// get enumerations from XPU for visu:	
GVL_APPLICATION.VisuPoolData.eTransportState                       := f_GetState   (GVL_XTS.XtsTransportState.State);
GVL_APPLICATION.VisuPoolData.eTransportResult                      := f_GetProgress(GVL_XTS.XtsTransportState.State);
GVL_APPLICATION.VisuPoolData.eXpuState                             := f_GetState   (GVL_XTS.XtsTransportState.XpuState.State);
GVL_APPLICATION.VisuPoolData.eXpuResult                            := f_GetProgress(GVL_XTS.XtsTransportState.XpuState.State);
GVL_APPLICATION.VisuPoolData.eXpuCheck                             := GVL_XTS.XtsTransportState.XpuState.Check;

// display xpu state and result in visu
// get strings and info
GVL_APPLICATION.VisuPoolData.sCaGroupState                         := TO_STRING(GVL_XTS.XtsTransportState.GroupInfo.CaGroupState);

GVL_APPLICATION.VisuPoolData.sTransportState                       := TO_STRING(GVL_APPLICATION.VisuPoolData.eTransportState);
GVL_APPLICATION.VisuPoolData.sTransportCheck                       := TO_STRING(GVL_XTS.XtsTransportState.Check);
GVL_APPLICATION.VisuPoolData.sTransportResult                      := TO_STRING(GVL_APPLICATION.VisuPoolData.eTransportResult);

GVL_APPLICATION.VisuPoolData.stXpuStrings.sXpuState                := TO_STRING(GVL_APPLICATION.VisuPoolData.eXpuState);
GVL_APPLICATION.VisuPoolData.stXpuStrings.sXpuResult               := TO_STRING(GVL_APPLICATION.VisuPoolData.eXpuResult);
GVL_APPLICATION.VisuPoolData.stXpuStrings.sXpuCyclicCheck          := TO_STRING(GVL_APPLICATION.VisuPoolData.eXpuCheck);

GVL_APPLICATION.VisuPoolData.stXpuStrings.sXpuOpMode               := TO_STRING(GVL_XTS.XtsTransportState.XpuInfo.OperationMode);
GVL_APPLICATION.VisuPoolData.stXpuStrings.sXpuMoverId_DetectionMode:= TO_STRING(GVL_XTS.XtsTransportState.XpuInfo.IdDetectionMode);
GVL_APPLICATION.VisuPoolData.stXpuStrings.sXpuMoverPosAssignement  := TO_STRING(GVL_XTS.XtsTransportState.XpuInfo.MoverPositionAssignement);
//---------------------------------------------------------------------------------------------------------------
// check the indices before access
//---------------------------------------------------------------------------------------------------------------
nMoverSelected       := SEL((nMoverSelected<1),                               nMoverSelected, 1);
nMoverSelected       := SEL((nMoverSelected>GVL_XTS_CONSTANTS.MAX_MOVER),     nMoverSelected, GVL_XTS_CONSTANTS.MAX_MOVER);

nStationSelected     := SEL((nStationSelected<1),                             nStationSelected, 1);
nStationSelected     := SEL((nStationSelected>GVL_XTS_CONSTANTS.MAX_STATION), nStationSelected, GVL_XTS_CONSTANTS.MAX_STATION);

nCollectorSelected   := SEL((nCollectorSelected<1),                           nCollectorSelected, 1);
nCollectorSelected   := SEL((nCollectorSelected>GVL_APPLICATION.MAX_PROCESS), nCollectorSelected, GVL_APPLICATION.MAX_PROCESS);

nInstanceSelected    := SEL((nInstanceSelected<1),                            nInstanceSelected, 1);
nInstanceSelected    := SEL((nInstanceSelected>GVL_APPLICATION.MAX_PROCESS),  nInstanceSelected, GVL_APPLICATION.MAX_PROCESS);
//---------------------------------------------------------------------------------------------------------------
// get indexed data
//---------------------------------------------------------------------------------------------------------------
GVL_APPLICATION.VisuPoolData.eMoverState        := f_GetState   (GVL_XTS.MoverState[nMoverSelected].State);
GVL_APPLICATION.VisuPoolData.eMoverResult       := f_GetProgress(GVL_XTS.MoverState[nMoverSelected].State);
GVL_APPLICATION.VisuPoolData.sMoverState        := TO_STRING(GVL_APPLICATION.VisuPoolData.eMoverState);
GVL_APPLICATION.VisuPoolData.sMoverResult       := TO_STRING(GVL_APPLICATION.VisuPoolData.eMoverResult);

GVL_APPLICATION.VisuPoolData.bStationEnable     := SEL((GVL_XTS.StationCtrl[nStationSelected].Cmd = E_STATION_CTRL.STATION_ENABLE),        FALSE, TRUE);
GVL_APPLICATION.VisuPoolData.bStationEnter      := SEL((GVL_XTS.StationCtrl[nStationSelected].Cmd = E_STATION_CTRL.STATION_MOVER_ENTER),   FALSE, TRUE);
GVL_APPLICATION.VisuPoolData.bStationStart      := SEL((GVL_XTS.StationCtrl[nStationSelected].Cmd = E_STATION_CTRL.STATION_PROCESS_START), FALSE, TRUE);
GVL_APPLICATION.VisuPoolData.bStationDone       := SEL((GVL_XTS.StationCtrl[nStationSelected].Cmd = E_STATION_CTRL.STATION_PROCESS_DONE),  FALSE, TRUE);
GVL_APPLICATION.VisuPoolData.bStationOut        := SEL((GVL_XTS.StationCtrl[nStationSelected].Cmd = E_STATION_CTRL.STATION_MOVER_OUT),     FALSE, TRUE);
GVL_APPLICATION.VisuPoolData.bStationGone       := SEL((GVL_XTS.StationCtrl[nStationSelected].Cmd = E_STATION_CTRL.STATION_MOVER_GONE),    FALSE, TRUE);

GVL_APPLICATION.VisuPoolData.sStationState      := TO_STRING(GVL_XTS.StationState[nStationSelected].State);
GVL_APPLICATION.VisuPoolData.sStationStateMask  := Tc2_Utilities.BYTE_TO_BINSTR(GVL_XTS.StationState[nStationSelected].nMask, 8);
GVL_APPLICATION.VisuPoolData.sStationCtrlMask   := Tc2_Utilities.BYTE_TO_BINSTR(GVL_XTS.StationCtrl[nStationSelected].nMask, 8);
//---------------------------------------------------------------------------------------------------------------
// Mover Selector
//---------------------------------------------------------------------------------------------------------------
GVL_APPLICATION.VisuPoolData.eSelectorState     := f_GetState   (GVL_XTS.MoverSelectorState.State.State);
GVL_APPLICATION.VisuPoolData.eSelectorResult    := f_GetProgress(GVL_XTS.MoverSelectorState.State.State);
GVL_APPLICATION.VisuPoolData.sSelectorState     := TO_STRING(GVL_APPLICATION.VisuPoolData.eSelectorState);
GVL_APPLICATION.VisuPoolData.sSelectorResult    := TO_STRING(GVL_APPLICATION.VisuPoolData.eSelectorResult);
//---------------------------------------------------------------------------------------------------------------
//---------------------------------------------------------------------------------------------------------------
//---------------------------------------------------------------------------------------------------------------

END_PROGRAM

// ---- APPLICATION/MAIN_APP.TcPOU
//---------------------------------------------------------------------------------------------------------------
//
//  HAUD 2026.10.25
//
//  - ExternControl
//
//    - this is the main switchboard
//
//    - Transport abstractions are called here:
//    --------------------------------------------
//    - top level transport abstractions
//      - Instances contain the required transport logic
//      - Instances control their assigned ProcessCollector
//      - Instances are controlled in timer based application
//
//    - mid level transport abstractions
//      - StationCollectors and by extension ProcessCollectors
//      - Collectors are for gathering states and routing commands to ST_STATION_CTRL/STATE
//      - Collectors are configured during startup
//
//---------------------------------------------------------------------------------------------------------------
PROGRAM MAIN_APP
VAR
  eInitXtsTransport   AT %I*    : E_PROGRESS;   // initialization from XtsTransport PLC
  eInit               AT %Q*    : E_PROGRESS;   // local startup transmitted to TowerControl

  idx                           : UINT;
  nProcess                      : E_INSTANCE;

  // message pipeline(s) handling
  eMtrState,
  eMsgState                     : E_MESSAGE_STATE;
  eMtrProgress,
  eMsgProgress                  : E_PROGRESS;
  stMsg                         : ST_Message;
  //-------------------------------------------------------------------------------------------------------------
  tIdleWriteMotion              : TIME := T#5S;
  tIdleWriteApplication         : TIME := T#5S;
  tIdleWriteMetric              : TIME := T#5S;
  tonIdleWriteMotion            : Tc2_Standard.TON;
  tonIdleWriteApplication       : Tc2_Standard.TON;
  tonIdleWriteMetric            : Tc2_Standard.TON;
  //-------------------------------------------------------------------------------------------------------------
END_VAR

//#################################################################################################################
// Local time; used for timestamps
//#################################################################################################################
GVL_MSG_XTS.fbLocalTime();
GVL_MSG_XTS.sLocalTime                                            := GVL_MSG_XTS.fbLocalTime.LocalTimeString;
GVL_MSG_XTS.dtLocalTime                                           := GVL_MSG_XTS.fbLocalTime.LocalTime;
//-----------------------------------------------------------------------------------------------------------------
//-----------------------------------------------------------------------------------------------------------------
// check for Initialisation from XtsTransport first
//  - wait for XtsTransport to be fully started up
//-----------------------------------------------------------------------------------------------------------------
IF NOT (eInitXtsTransport = E_PROGRESS.PROGRESS_DONE) THEN eInit  := E_PROGRESS.PROGRESS_INVALID; RETURN; END_IF
//-----------------------------------------------------------------------------------------------------------------
//-----------------------------------------------------------------------------------------------------------------
// initialization for:
//  - configuring processes
//  - starting up of processes
//  - cross checking with the rest of your application
//-----------------------------------------------------------------------------------------------------------------
CASE eInit
OF
  E_PROGRESS.PROGRESS_INVALID:
    GVL_MSG_XTS.MetricsMessageCtrl.Cmd            := E_MESSAGE_CTRL.MSG_CTRL_INIT;
    eInit                                         := E_PROGRESS.PROGRESS_INIT;

  E_PROGRESS.PROGRESS_INIT:
    // init processes
    eInit                                         := E_PROGRESS.PROGRESS_BUSY;
    //-----------------------------------------------------------------------------
    //#############################################################################
    //-----------------------------------------------------------------------------
    GVL_APPLICATION.ProcessCollector[DISTRIBUTOR_INFEED].ProcessId            := DISTRIBUTOR_INFEED;
    GVL_APPLICATION.ProcessCollector[DISTRIBUTOR_INFEED].StationFirst         :=   142;
    GVL_APPLICATION.ProcessCollector[DISTRIBUTOR_INFEED].StationLast          :=   142;
    //-----------------------------------------------------------------------------
    GVL_APPLICATION.InstanceDistributorInfeed.ProcessId                       := DISTRIBUTOR_INFEED;
    GVL_APPLICATION.InstanceDistributorInfeed.ProcessTarget                   := PROCESS_INFEED;
    GVL_APPLICATION.InstanceDistributorInfeed.CheckPositionStart              :=  4500.0;
    GVL_APPLICATION.InstanceDistributorInfeed.CheckPositionEnd                :=  5600.0;
    //-----------------------------------------------------------------------------
    GVL_APPLICATION.InstanceDistributorInfeed.CollectorInterface              :=   GVL_APPLICATION.ItfProcessCollector;
    GVL_APPLICATION.InstanceDistributorInfeed.ProcessLinkedLists              :=   GVL_APPLICATION.ItfProcessList;
    GVL_APPLICATION.InstanceDistributorInfeed.InstanceCtrl                    REF= GVL_APPLICATION.InstanceCtrl;
    GVL_APPLICATION.InstanceDistributorInfeed.InstanceState                   REF= GVL_APPLICATION.InstanceState;
    GVL_APPLICATION.InstanceDistributorInfeed.MessageLevel                    :=   E_MessageType.eMessageError;

    //-----------------------------------------------------------------------------
    //#############################################################################
    //-----------------------------------------------------------------------------
    GVL_APPLICATION.ProcessCollector[PROCESS_INFEED].ProcessId                := PROCESS_INFEED;
    GVL_APPLICATION.ProcessCollector[PROCESS_INFEED].StationFirst             :=    20;
    GVL_APPLICATION.ProcessCollector[PROCESS_INFEED].StationLast              :=    35;
    //-----------------------------------------------------------------------------
    GVL_APPLICATION.InstanceInfeed.ProcessId                                  := PROCESS_INFEED;
    GVL_APPLICATION.InstanceInfeed.ProcessTarget                              := CONTINUOUS_CLEAN;
    GVL_APPLICATION.InstanceInfeed.CheckPositionStart                         :=  9750.0;
    GVL_APPLICATION.InstanceInfeed.CheckPositionEnd                           := 12100.0;
    //-----------------------------------------------------------------------------
    GVL_APPLICATION.InstanceInfeed.CollectorInterface                         :=   GVL_APPLICATION.ItfProcessCollector;
    GVL_APPLICATION.InstanceInfeed.ProcessLinkedLists                         :=   GVL_APPLICATION.ItfProcessList;
    GVL_APPLICATION.InstanceInfeed.InstanceCtrl                               REF= GVL_APPLICATION.InstanceCtrl;
    GVL_APPLICATION.InstanceInfeed.InstanceState                              REF= GVL_APPLICATION.InstanceState;
    GVL_APPLICATION.InstanceInfeed.MessageLevel                               :=   E_MessageType.eMessageError;

    //-----------------------------------------------------------------------------
    //#############################################################################
    //-----------------------------------------------------------------------------
    GVL_APPLICATION.ProcessCollector[CONTINUOUS_CLEAN].ProcessId              := CONTINUOUS_CLEAN;
    GVL_APPLICATION.ProcessCollector[CONTINUOUS_CLEAN].StationFirst           :=    37;
    GVL_APPLICATION.ProcessCollector[CONTINUOUS_CLEAN].StationLast            :=    37;
    //-----------------------------------------------------------------------------
    GVL_APPLICATION.InstanceCleaner.ProcessId                                 := CONTINUOUS_CLEAN;
    GVL_APPLICATION.InstanceCleaner.ProcessTarget                             := CONTINUOUS_SCAN;
    GVL_APPLICATION.InstanceCleaner.CheckPositionStart                        := 12850.0;
    GVL_APPLICATION.InstanceCleaner.CheckPositionEnd                          := 13000.0;
    //-----------------------------------------------------------------------------
    GVL_APPLICATION.InstanceCleaner.CollectorInterface                        :=   GVL_APPLICATION.ItfProcessCollector;
    GVL_APPLICATION.InstanceCleaner.ProcessLinkedLists                        :=   GVL_APPLICATION.ItfProcessList;
    GVL_APPLICATION.InstanceCleaner.InstanceCtrl                              REF= GVL_APPLICATION.InstanceCtrl;
    GVL_APPLICATION.InstanceCleaner.InstanceState                             REF= GVL_APPLICATION.InstanceState;

    //-----------------------------------------------------------------------------
    //#############################################################################
    //-----------------------------------------------------------------------------
    GVL_APPLICATION.ProcessCollector[CONTINUOUS_SCAN].ProcessId               := CONTINUOUS_SCAN;
    GVL_APPLICATION.ProcessCollector[CONTINUOUS_SCAN].StationFirst            :=    38;
    GVL_APPLICATION.ProcessCollector[CONTINUOUS_SCAN].StationLast             :=    38;
    //-----------------------------------------------------------------------------
    GVL_APPLICATION.InstanceScanner.ProcessId                                 := CONTINUOUS_SCAN;
    GVL_APPLICATION.InstanceScanner.ProcessTarget                             := CONTINUOUS_CAMERA;
    GVL_APPLICATION.InstanceScanner.CheckPositionStart                        := 13900.0;
    GVL_APPLICATION.InstanceScanner.CheckPositionEnd                          := 14100.0;
    //-----------------------------------------------------------------------------
    GVL_APPLICATION.InstanceScanner.CollectorInterface                        :=   GVL_APPLICATION.ItfProcessCollector;
    GVL_APPLICATION.InstanceScanner.ProcessLinkedLists                        :=   GVL_APPLICATION.ItfProcessList;
    GVL_APPLICATION.InstanceScanner.InstanceCtrl                              REF= GVL_APPLICATION.InstanceCtrl;
    GVL_APPLICATION.InstanceScanner.InstanceState                             REF= GVL_APPLICATION.InstanceState;

    //-----------------------------------------------------------------------------
    //#############################################################################
    //-----------------------------------------------------------------------------
    GVL_APPLICATION.ProcessCollector[CONTINUOUS_CAMERA].ProcessId             := CONTINUOUS_CAMERA;
    GVL_APPLICATION.ProcessCollector[CONTINUOUS_CAMERA].StationFirst          :=    39;
    GVL_APPLICATION.ProcessCollector[CONTINUOUS_CAMERA].StationLast           :=    39;
    //-----------------------------------------------------------------------------
    GVL_APPLICATION.InstanceCamera.ProcessId                                  := CONTINUOUS_CAMERA;
    GVL_APPLICATION.InstanceCamera.ProcessTarget                              := DISTRIBUTOR_ASSEMBLY_01;
    GVL_APPLICATION.InstanceCamera.CheckPositionStart                         := 14200.0;
    GVL_APPLICATION.InstanceCamera.CheckPositionEnd                           := 14400.0;
    //-----------------------------------------------------------------------------
    GVL_APPLICATION.InstanceCamera.CollectorInterface                         :=   GVL_APPLICATION.ItfProcessCollector;
    GVL_APPLICATION.InstanceCamera.ProcessLinkedLists                         :=   GVL_APPLICATION.ItfProcessList;
    GVL_APPLICATION.InstanceCamera.InstanceCtrl                               REF= GVL_APPLICATION.InstanceCtrl;
    GVL_APPLICATION.InstanceCamera.InstanceState                              REF= GVL_APPLICATION.InstanceState;

    //-----------------------------------------------------------------------------
    //#############################################################################
    //-----------------------------------------------------------------------------
    GVL_APPLICATION.ProcessCollector[DISTRIBUTOR_ASSEMBLY_01].ProcessId       := DISTRIBUTOR_ASSEMBLY_01;
    GVL_APPLICATION.ProcessCollector[DISTRIBUTOR_ASSEMBLY_01].StationFirst    :=    40;
    GVL_APPLICATION.ProcessCollector[DISTRIBUTOR_ASSEMBLY_01].StationLast     :=    40;
    //-----------------------------------------------------------------------------
    GVL_APPLICATION.InstanceDistributorAssembly_01.ProcessId                  := DISTRIBUTOR_ASSEMBLY_01;
    GVL_APPLICATION.InstanceDistributorAssembly_01.ProcessTarget              := PROCESS_ASSEMBLY_01;
    GVL_APPLICATION.InstanceDistributorAssembly_01.CheckPositionStart         := 14400.0;
    GVL_APPLICATION.InstanceDistributorAssembly_01.CheckPositionEnd           := 17500.0;
    //-----------------------------------------------------------------------------
    GVL_APPLICATION.InstanceDistributorAssembly_01.CollectorInterface         :=   GVL_APPLICATION.ItfProcessCollector;
    GVL_APPLICATION.InstanceDistributorAssembly_01.ProcessLinkedLists         :=   GVL_APPLICATION.ItfProcessList;
    GVL_APPLICATION.InstanceDistributorAssembly_01.InstanceCtrl               REF= GVL_APPLICATION.InstanceCtrl;
    GVL_APPLICATION.InstanceDistributorAssembly_01.InstanceState              REF= GVL_APPLICATION.InstanceState;

    //-----------------------------------------------------------------------------
    //#############################################################################
    //-----------------------------------------------------------------------------
    GVL_APPLICATION.ProcessCollector[PROCESS_ASSEMBLY_01].ProcessId           := PROCESS_ASSEMBLY_01;
    GVL_APPLICATION.ProcessCollector[PROCESS_ASSEMBLY_01].StationFirst        :=    41;
    GVL_APPLICATION.ProcessCollector[PROCESS_ASSEMBLY_01].StationLast         :=    56;
    //-----------------------------------------------------------------------------
    GVL_APPLICATION.InstanceAssembly_01.ProcessId                             := PROCESS_ASSEMBLY_01;
    GVL_APPLICATION.InstanceAssembly_01.ProcessTarget                         := DISTRIBUTOR_ASSEMBLY_02;
    GVL_APPLICATION.InstanceAssembly_01.CheckPositionStart                    := 14400.0;
    GVL_APPLICATION.InstanceAssembly_01.CheckPositionEnd                      := 17500.0;
    //-----------------------------------------------------------------------------
    GVL_APPLICATION.InstanceAssembly_01.CollectorInterface                    :=   GVL_APPLICATION.ItfProcessCollector;
    GVL_APPLICATION.InstanceAssembly_01.ProcessLinkedLists                    :=   GVL_APPLICATION.ItfProcessList;
    GVL_APPLICATION.InstanceAssembly_01.InstanceCtrl                          REF= GVL_APPLICATION.InstanceCtrl;
    GVL_APPLICATION.InstanceAssembly_01.InstanceState                         REF= GVL_APPLICATION.InstanceState;

    //-----------------------------------------------------------------------------
    //#############################################################################
    //-----------------------------------------------------------------------------
    GVL_APPLICATION.ProcessCollector[DISTRIBUTOR_ASSEMBLY_02].ProcessId       := DISTRIBUTOR_ASSEMBLY_02;
    GVL_APPLICATION.ProcessCollector[DISTRIBUTOR_ASSEMBLY_02].StationFirst    :=    57;
    GVL_APPLICATION.ProcessCollector[DISTRIBUTOR_ASSEMBLY_02].StationLast     :=    57;
    //-----------------------------------------------------------------------------
    GVL_APPLICATION.InstanceDistributorAssembly_02.ProcessId                  := DISTRIBUTOR_ASSEMBLY_02;
    GVL_APPLICATION.InstanceDistributorAssembly_02.ProcessTarget              := PROCESS_ASSEMBLY_02;
    GVL_APPLICATION.InstanceDistributorAssembly_02.CheckPositionStart         := 17500.0;
    GVL_APPLICATION.InstanceDistributorAssembly_02.CheckPositionEnd           := 18100.0;
    //-----------------------------------------------------------------------------
    GVL_APPLICATION.InstanceDistributorAssembly_02.CollectorInterface         :=   GVL_APPLICATION.ItfProcessCollector;
    GVL_APPLICATION.InstanceDistributorAssembly_02.ProcessLinkedLists         :=   GVL_APPLICATION.ItfProcessList;
    GVL_APPLICATION.InstanceDistributorAssembly_02.InstanceCtrl               REF= GVL_APPLICATION.InstanceCtrl;
    GVL_APPLICATION.InstanceDistributorAssembly_02.InstanceState              REF= GVL_APPLICATION.InstanceState;

    //-----------------------------------------------------------------------------
    //#############################################################################
    //-----------------------------------------------------------------------------
    GVL_APPLICATION.ProcessCollector[PROCESS_ASSEMBLY_02].ProcessId           := PROCESS_ASSEMBLY_02;
    GVL_APPLICATION.ProcessCollector[PROCESS_ASSEMBLY_02].StationFirst        :=    58;
    GVL_APPLICATION.ProcessCollector[PROCESS_ASSEMBLY_02].StationLast         :=    67;
    //-----------------------------------------------------------------------------
    GVL_APPLICATION.InstanceAssembly_02.ProcessId                             := PROCESS_ASSEMBLY_02;
    GVL_APPLICATION.InstanceAssembly_02.ProcessTarget                         := DISTRIBUTOR_ASSEMBLY_TEST;
    GVL_APPLICATION.InstanceAssembly_02.CheckPositionStart                    := 19400.0;
    GVL_APPLICATION.InstanceAssembly_02.CheckPositionEnd                      := 20750.0;
    //-----------------------------------------------------------------------------
    GVL_APPLICATION.InstanceAssembly_02.CollectorInterface                    :=   GVL_APPLICATION.ItfProcessCollector;
    GVL_APPLICATION.InstanceAssembly_02.ProcessLinkedLists                    :=   GVL_APPLICATION.ItfProcessList;
    GVL_APPLICATION.InstanceAssembly_02.InstanceCtrl                          REF= GVL_APPLICATION.InstanceCtrl;
    GVL_APPLICATION.InstanceAssembly_02.InstanceState                         REF= GVL_APPLICATION.InstanceState;

    //-----------------------------------------------------------------------------
    //#############################################################################
    //-----------------------------------------------------------------------------
    GVL_APPLICATION.ProcessCollector[DISTRIBUTOR_ASSEMBLY_TEST].ProcessId     := DISTRIBUTOR_ASSEMBLY_TEST;
    GVL_APPLICATION.ProcessCollector[DISTRIBUTOR_ASSEMBLY_TEST].StationFirst  :=    70;
    GVL_APPLICATION.ProcessCollector[DISTRIBUTOR_ASSEMBLY_TEST].StationLast   :=    70;
    //-----------------------------------------------------------------------------
    GVL_APPLICATION.InstanceDistributorAssemblyTest.ProcessId                 := DISTRIBUTOR_ASSEMBLY_TEST;
    GVL_APPLICATION.InstanceDistributorAssemblyTest.ProcessTarget             := PROCESS_ASSEMBLY_TEST;
    GVL_APPLICATION.InstanceDistributorAssemblyTest.CheckPositionStart        := 20600.0;
    GVL_APPLICATION.InstanceDistributorAssemblyTest.CheckPositionEnd          := 21400.0;
    //-----------------------------------------------------------------------------
    GVL_APPLICATION.InstanceDistributorAssemblyTest.CollectorInterface        :=   GVL_APPLICATION.ItfProcessCollector;
    GVL_APPLICATION.InstanceDistributorAssemblyTest.ProcessLinkedLists        :=   GVL_APPLICATION.ItfProcessList;
    GVL_APPLICATION.InstanceDistributorAssemblyTest.InstanceCtrl              REF= GVL_APPLICATION.InstanceCtrl;
    GVL_APPLICATION.InstanceDistributorAssemblyTest.InstanceState             REF= GVL_APPLICATION.InstanceState;

    //-----------------------------------------------------------------------------
    //#############################################################################
    //-----------------------------------------------------------------------------
    GVL_APPLICATION.ProcessCollector[PROCESS_ASSEMBLY_TEST].ProcessId         := PROCESS_ASSEMBLY_TEST;
    GVL_APPLICATION.ProcessCollector[PROCESS_ASSEMBLY_TEST].StationFirst      :=    71;
    GVL_APPLICATION.ProcessCollector[PROCESS_ASSEMBLY_TEST].StationLast       :=    86;
    //-----------------------------------------------------------------------------
    GVL_APPLICATION.InstanceAssemblyTest.ProcessId                            := PROCESS_ASSEMBLY_TEST;
    GVL_APPLICATION.InstanceAssemblyTest.ProcessTarget                        := DISTRIBUTOR_CAMERA;
    GVL_APPLICATION.InstanceAssemblyTest.CheckPositionStart                   := 21400.0;
    GVL_APPLICATION.InstanceAssemblyTest.CheckPositionEnd                     := 23000.0;
    //-----------------------------------------------------------------------------
    GVL_APPLICATION.InstanceAssemblyTest.CollectorInterface                   :=   GVL_APPLICATION.ItfProcessCollector;
    GVL_APPLICATION.InstanceAssemblyTest.ProcessLinkedLists                   :=   GVL_APPLICATION.ItfProcessList;
    GVL_APPLICATION.InstanceAssemblyTest.InstanceCtrl                         REF= GVL_APPLICATION.InstanceCtrl;
    GVL_APPLICATION.InstanceAssemblyTest.InstanceState                        REF= GVL_APPLICATION.InstanceState;

    //-----------------------------------------------------------------------------
    //#############################################################################
    //-----------------------------------------------------------------------------
    GVL_APPLICATION.ProcessCollector[DISTRIBUTOR_CAMERA].ProcessId            := DISTRIBUTOR_CAMERA;
    GVL_APPLICATION.ProcessCollector[DISTRIBUTOR_CAMERA].StationFirst         :=    91;
    GVL_APPLICATION.ProcessCollector[DISTRIBUTOR_CAMERA].StationLast          :=    91;
    //-----------------------------------------------------------------------------
    GVL_APPLICATION.InstanceAssemblyCameraInfeed.ProcessId                    := DISTRIBUTOR_CAMERA;
    GVL_APPLICATION.InstanceAssemblyCameraInfeed.ProcessTarget                := CONTINUOUS_ASSEMBLY_CAMERA;
    GVL_APPLICATION.InstanceAssemblyCameraInfeed.CheckPositionStart           := 22800.0;
    GVL_APPLICATION.InstanceAssemblyCameraInfeed.CheckPositionEnd             := 23500.0;
    //-----------------------------------------------------------------------------
    GVL_APPLICATION.InstanceAssemblyCameraInfeed.CollectorInterface           :=   GVL_APPLICATION.ItfProcessCollector;
    GVL_APPLICATION.InstanceAssemblyCameraInfeed.ProcessLinkedLists           :=   GVL_APPLICATION.ItfProcessList;
    GVL_APPLICATION.InstanceAssemblyCameraInfeed.InstanceCtrl                 REF= GVL_APPLICATION.InstanceCtrl;
    GVL_APPLICATION.InstanceAssemblyCameraInfeed.InstanceState                REF= GVL_APPLICATION.InstanceState;

    //-----------------------------------------------------------------------------
    //#############################################################################
    //-----------------------------------------------------------------------------
    GVL_APPLICATION.ProcessCollector[CONTINUOUS_ASSEMBLY_CAMERA].ProcessId    := CONTINUOUS_ASSEMBLY_CAMERA;
    GVL_APPLICATION.ProcessCollector[CONTINUOUS_ASSEMBLY_CAMERA].StationFirst :=    95;
    GVL_APPLICATION.ProcessCollector[CONTINUOUS_ASSEMBLY_CAMERA].StationLast  :=    95;
    //-----------------------------------------------------------------------------
    GVL_APPLICATION.InstanceAssemblyCameraOutfeed.ProcessId                   := CONTINUOUS_ASSEMBLY_CAMERA;
    GVL_APPLICATION.InstanceAssemblyCameraOutfeed.ProcessTarget               := DISTRIBUTOR_OUTFEED;
    GVL_APPLICATION.InstanceAssemblyCameraOutfeed.CheckPositionStart          := 24000.0;
    GVL_APPLICATION.InstanceAssemblyCameraOutfeed.CheckPositionEnd            := 24100.0;
    //-----------------------------------------------------------------------------
    GVL_APPLICATION.InstanceAssemblyCameraOutfeed.CollectorInterface          :=   GVL_APPLICATION.ItfProcessCollector;
    GVL_APPLICATION.InstanceAssemblyCameraOutfeed.ProcessLinkedLists          :=   GVL_APPLICATION.ItfProcessList;
    GVL_APPLICATION.InstanceAssemblyCameraOutfeed.InstanceCtrl                REF= GVL_APPLICATION.InstanceCtrl;
    GVL_APPLICATION.InstanceAssemblyCameraOutfeed.InstanceState               REF= GVL_APPLICATION.InstanceState;

    //-----------------------------------------------------------------------------
    //#############################################################################
    //-----------------------------------------------------------------------------
    GVL_APPLICATION.ProcessCollector[DISTRIBUTOR_OUTFEED].ProcessId           := DISTRIBUTOR_OUTFEED;
    GVL_APPLICATION.ProcessCollector[DISTRIBUTOR_OUTFEED].StationFirst        :=   119;
    GVL_APPLICATION.ProcessCollector[DISTRIBUTOR_OUTFEED].StationLast         :=   119;
    //-----------------------------------------------------------------------------
    GVL_APPLICATION.InstanceDistributorOutfeed.ProcessId                      := DISTRIBUTOR_OUTFEED;
    GVL_APPLICATION.InstanceDistributorOutfeed.ProcessTarget                  := PROCESS_OUTFEED;
    GVL_APPLICATION.InstanceDistributorOutfeed.CheckPositionStart             := 24000.0;
    GVL_APPLICATION.InstanceDistributorOutfeed.CheckPositionEnd               := 27500.0;
    //-----------------------------------------------------------------------------
    GVL_APPLICATION.InstanceDistributorOutfeed.CollectorInterface             :=   GVL_APPLICATION.ItfProcessCollector;
    GVL_APPLICATION.InstanceDistributorOutfeed.ProcessLinkedLists             :=   GVL_APPLICATION.ItfProcessList;
    GVL_APPLICATION.InstanceDistributorOutfeed.InstanceCtrl                   REF= GVL_APPLICATION.InstanceCtrl;
    GVL_APPLICATION.InstanceDistributorOutfeed.InstanceState                  REF= GVL_APPLICATION.InstanceState;

    //-----------------------------------------------------------------------------
    //#############################################################################
    //-----------------------------------------------------------------------------
    GVL_APPLICATION.ProcessCollector[PROCESS_OUTFEED].ProcessId               := PROCESS_OUTFEED;
    GVL_APPLICATION.ProcessCollector[PROCESS_OUTFEED].StationFirst            :=   120;
    GVL_APPLICATION.ProcessCollector[PROCESS_OUTFEED].StationLast             :=   133;
    //-----------------------------------------------------------------------------
    GVL_APPLICATION.InstanceOutfeed.ProcessId                                 := PROCESS_OUTFEED;
    GVL_APPLICATION.InstanceOutfeed.ProcessTarget                             := DISTRIBUTOR_WPC_CLEAN;
    GVL_APPLICATION.InstanceOutfeed.CheckPositionStart                        := 24500.0;
    GVL_APPLICATION.InstanceOutfeed.CheckPositionEnd                          := 27500.0;
    //-----------------------------------------------------------------------------
    GVL_APPLICATION.InstanceOutfeed.CollectorInterface                        :=   GVL_APPLICATION.ItfProcessCollector;
    GVL_APPLICATION.InstanceOutfeed.ProcessLinkedLists                        :=   GVL_APPLICATION.ItfProcessList;
    GVL_APPLICATION.InstanceOutfeed.InstanceCtrl                              REF= GVL_APPLICATION.InstanceCtrl;
    GVL_APPLICATION.InstanceOutfeed.InstanceState                             REF= GVL_APPLICATION.InstanceState;

    //-----------------------------------------------------------------------------
    //#############################################################################
    //-----------------------------------------------------------------------------
    GVL_APPLICATION.ProcessCollector[DISTRIBUTOR_WPC_CLEAN].ProcessId         := DISTRIBUTOR_WPC_CLEAN;
    GVL_APPLICATION.ProcessCollector[DISTRIBUTOR_WPC_CLEAN].StationFirst      :=   140;
    GVL_APPLICATION.ProcessCollector[DISTRIBUTOR_WPC_CLEAN].StationLast       :=   140;
    //-----------------------------------------------------------------------------
    GVL_APPLICATION.InstanceDistributorWpcClean.ProcessId                     := DISTRIBUTOR_WPC_CLEAN;
    GVL_APPLICATION.InstanceDistributorWpcClean.ProcessTarget                 := CONTINUOUS_WPC_CLEAN;
    GVL_APPLICATION.InstanceDistributorWpcClean.CheckPositionStart            := 27970.0;
    GVL_APPLICATION.InstanceDistributorWpcClean.CheckPositionEnd              :=  1250.0;
    //-----------------------------------------------------------------------------
    GVL_APPLICATION.InstanceDistributorWpcClean.CollectorInterface            :=   GVL_APPLICATION.ItfProcessCollector;
    GVL_APPLICATION.InstanceDistributorWpcClean.ProcessLinkedLists            :=   GVL_APPLICATION.ItfProcessList;
    GVL_APPLICATION.InstanceDistributorWpcClean.InstanceCtrl                  REF= GVL_APPLICATION.InstanceCtrl;
    GVL_APPLICATION.InstanceDistributorWpcClean.InstanceState                 REF= GVL_APPLICATION.InstanceState;

    //-----------------------------------------------------------------------------
    //#############################################################################
    //-----------------------------------------------------------------------------
    GVL_APPLICATION.ProcessCollector[CONTINUOUS_WPC_CLEAN].ProcessId          := CONTINUOUS_WPC_CLEAN;
    GVL_APPLICATION.ProcessCollector[CONTINUOUS_WPC_CLEAN].StationFirst       :=   141;
    GVL_APPLICATION.ProcessCollector[CONTINUOUS_WPC_CLEAN].StationLast        :=   141;
    //-----------------------------------------------------------------------------
    GVL_APPLICATION.InstanceWpcClean.ProcessId                                := CONTINUOUS_WPC_CLEAN;
    GVL_APPLICATION.InstanceWpcClean.ProcessTarget                            := DISTRIBUTOR_INFEED;
    GVL_APPLICATION.InstanceWpcClean.CheckPositionStart                       :=  3950.0;
    GVL_APPLICATION.InstanceWpcClean.CheckPositionEnd                         :=  4100.0;
    //-----------------------------------------------------------------------------
    GVL_APPLICATION.InstanceWpcClean.CollectorInterface                       :=   GVL_APPLICATION.ItfProcessCollector;
    GVL_APPLICATION.InstanceWpcClean.ProcessLinkedLists                       :=   GVL_APPLICATION.ItfProcessList;
    GVL_APPLICATION.InstanceWpcClean.InstanceCtrl                             REF= GVL_APPLICATION.InstanceCtrl;
    GVL_APPLICATION.InstanceWpcClean.InstanceState                            REF= GVL_APPLICATION.InstanceState;


  E_PROGRESS.PROGRESS_BUSY:
    // init the conductor
    GVL_APPLICATION.ConductorCtrl.Cmd             := E_INSTANCE_CMD.INIT;
    // init the instances
    idx                                           := 1;
    memset(ADR(GVL_APPLICATION.InstanceCtrl), 0, SIZEOF(GVL_APPLICATION.InstanceCtrl));
    eInit                                         := E_PROGRESS.PROGRESS_PREPARE;

  E_PROGRESS.PROGRESS_PREPARE:
    GVL_APPLICATION.InstanceCtrl[idx].Cmd         := E_INSTANCE_CMD.INIT;

    IF (GVL_APPLICATION.InstanceState[idx].ProcessState   = E_INSTANCE_STATE.DISABLED)
    THEN
      IF (GVL_APPLICATION.InstanceState[idx].ProcessProgress = E_PROGRESS.PROGRESS_BUSY)
      THEN
        GVL_APPLICATION.InstanceCtrl[idx].Cmd     := E_INSTANCE_CMD.DISABLE;
        eInit                                     := E_PROGRESS.PROGRESS_STARTUP;
      END_IF
    END_IF


  E_PROGRESS.PROGRESS_STARTUP:
    IF NOT (idx < GVL_APPLICATION.MAX_PROCESS)
    THEN
      eInit                                       := E_PROGRESS.PROGRESS_CHECK;
    ELSE
      idx                                         := idx + 1;
      eInit                                       := E_PROGRESS.PROGRESS_PREPARE;
    END_IF

  E_PROGRESS.PROGRESS_CHECK:
    GVL_APPLICATION.ConductorCtrl.Cmd             := E_INSTANCE_CMD.ENABLE;
    eInit                                         := E_PROGRESS.PROGRESS_OCCUPIED;

  E_PROGRESS.PROGRESS_OCCUPIED:
    eInit                                         := E_PROGRESS.PROGRESS_WORKING;

  E_PROGRESS.PROGRESS_WORKING:
    eInit                                         := E_PROGRESS.PROGRESS_DONE;
END_CASE
//-----------------------------------------------------------------------------------------------------------------
//-----------------------------------------------------------------------------------------------------------------
//-----------------------------------------------------------------------------------------------------------------
//-----------------------------------------------------------------------------------------------------------------
// /assign dataflow
//-----------------------------------------------------------------------------------------------------------------
//-----------------------------------------------------------------------------------------------------------------
//  - The YardMaster
//-----------------------------------------------------------------------------------------------------------------
GVL_APPLICATION.YardMaster.Ctrl                               REF= GVL_APPLICATION.YardControl;
GVL_APPLICATION.YardMaster.State                              REF= GVL_APPLICATION.YardState;

GVL_APPLICATION.YardMaster.XtsTransportCtrl                   REF= GVL_XTS.XtsTransportCtrl;
GVL_APPLICATION.YardMaster.XtsTransportState                  REF= GVL_XTS.XtsTransportState;

GVL_APPLICATION.YardMaster.CollectorInterfaces                :=   GVL_APPLICATION.ItfProcessCollector;
GVL_APPLICATION.YardMaster.TicketList                         :=   GVL_APPLICATION.TicketList;
GVL_APPLICATION.YardMaster();
//-----------------------------------------------------------------------------------------------------------------
//  - ProcessCollectors
//-----------------------------------------------------------------------------------------------------------------
FOR nProcess := 1 TO MAX_PROCESS
DO
  GVL_APPLICATION.ItfProcessList[nProcess]                    :=   GVL_APPLICATION.ProcessList[nProcess];
  GVL_APPLICATION.ItfProcessCollector[nProcess]               :=   GVL_APPLICATION.ProcessCollector[nProcess];

  GVL_APPLICATION.ProcessCollector[nProcess].MessageLevel     :=   GVL_MSG_XTS.MessageLevelProcess[nProcess];
  GVL_APPLICATION.ProcessCollector[nProcess].MoverInfo        REF= GVL_XTS.MoverInfo;
  GVL_APPLICATION.ProcessCollector[nProcess].StationCtrl      REF= GVL_XTS.StationCtrl;
  GVL_APPLICATION.ProcessCollector[nProcess].StationState     REF= GVL_XTS.StationState;
  GVL_APPLICATION.ProcessCollector[nProcess].Cycle();
END_FOR
//-----------------------------------------------------------------------------------------------------------------
//-----------------------------------------------------------------------------------------------------------------
// cyclic TicketList as inbox
//-----------------------------------------------------------------------------------------------------------------
//-----------------------------------------------------------------------------------------------------------------
GVL_APPLICATION.TicketControl.ItfList                         :=   GVL_APPLICATION.TicketList;
GVL_APPLICATION.TicketControl.Ctrl                            REF= GVL_APPLICATION.TicketListControl;
GVL_APPLICATION.TicketControl.State                           REF= GVL_APPLICATION.TicketListState;
GVL_APPLICATION.TicketControl.NodeDataInput                   REF= GVL_APPLICATION.TicketListDataInput;
GVL_APPLICATION.TicketControl.NodeDataOutput                  REF= GVL_APPLICATION.TicketListDataOutput;
GVL_APPLICATION.TicketControl();
//-----------------------------------------------------------------------------------------------------------------
//-----------------------------------------------------------------------------------------------------------------
// Conductor
//-----------------------------------------------------------------------------------------------------------------
//-----------------------------------------------------------------------------------------------------------------
GVL_APPLICATION.ProcessConductor.ProcessLinkedLists           :=   GVL_APPLICATION.ItfProcessList;
GVL_APPLICATION.ProcessConductor.TicketLinkedList             :=   GVL_APPLICATION.TicketList;
GVL_APPLICATION.ProcessConductor.Ctrl                         REF= GVL_APPLICATION.ConductorCtrl;
GVL_APPLICATION.ProcessConductor.State                        REF= GVL_APPLICATION.ConductorState;
GVL_APPLICATION.ProcessConductor();
//-----------------------------------------------------------------------------------------------------------------
//-----------------------------------------------------------------------------------------------------------------
// Instance calls
//-----------------------------------------------------------------------------------------------------------------
//-----------------------------------------------------------------------------------------------------------------
GVL_APPLICATION.InstanceWpcClean();
GVL_APPLICATION.InstanceDistributorWpcClean();
GVL_APPLICATION.InstanceOutfeed();
GVL_APPLICATION.InstanceDistributorOutfeed();
GVL_APPLICATION.InstanceAssemblyCameraOutfeed();
GVL_APPLICATION.InstanceAssemblyCameraInfeed();
GVL_APPLICATION.InstanceAssemblyTest();
GVL_APPLICATION.InstanceDistributorAssemblyTest();
GVL_APPLICATION.InstanceAssembly_02();
GVL_APPLICATION.InstanceDistributorAssembly_02();
GVL_APPLICATION.InstanceAssembly_01();
GVL_APPLICATION.InstanceDistributorAssembly_01();
GVL_APPLICATION.InstanceCamera();
GVL_APPLICATION.InstanceScanner();
GVL_APPLICATION.InstanceCleaner();
GVL_APPLICATION.InstanceInfeed();
GVL_APPLICATION.InstanceDistributorInfeed();
//-----------------------------------------------------------------------------------------------------------------
//-----------------------------------------------------------------------------------------------------------------
//#################################################################################################################
//  /logging
//    - all life is problem solving
//#################################################################################################################
GVL_MSG_XTS.TransportMessageData.Ctrl               REF= GVL_MSG_XTS.TransportMessageCtrl;
GVL_MSG_XTS.TransportMessageData.State              REF= GVL_MSG_XTS.TransportMessageState;
GVL_MSG_XTS.TransportMessageData.MessageIndex       REF= GVL_MSG_XTS.MessageTransportIndex;
GVL_MSG_XTS.TransportMessageData.ErrorIndex         REF= GVL_MSG_XTS.MessageTransportError;
GVL_MSG_XTS.TransportMessageData.DirRoot            :=   ADR(GVL_MSG_XTS.LOG_DIR);
GVL_MSG_XTS.TransportMessageData.FileRoot           :=   ADR(GVL_MSG_XTS.LOG_FILE);
GVL_MSG_XTS.TransportMessageData.MsgList            :=   ADR(GVL_MSG_XTS.TransportMessages);
GVL_MSG_XTS.TransportMessageData.LocalTime          :=   ADR(GVL_MSG_XTS.dtLocalTime);
GVL_MSG_XTS.TransportMessageData();
eMsgState                                       :=   f_GetState   (GVL_MSG_XTS.TransportMessageState.State);
eMsgProgress                                    :=   f_GetProgress(GVL_MSG_XTS.TransportMessageState.State);

CASE eMsgState
OF
  E_MESSAGE_STATE.MSG_STATE_NULL:
    CASE eMsgProgress
    OF
      E_PROGRESS.PROGRESS_INVALID,
      E_PROGRESS.PROGRESS_DONE:
        IF (GVL_MSG_XTS.MessageTransportIndex > GVL_MSG_XTS.MAX_MESSAGE/101) OR
           (GVL_MSG_XTS.MessageTransportError > 0)
        THEN
          GVL_MSG_XTS.TransportMessageCtrl.Cmd      := E_MESSAGE_CTRL.MSG_CTRL_WRITE;
        ELSE
          tonIdleWriteMotion(IN := TRUE, PT:= tIdleWriteMotion);
          IF (tonIdleWriteMotion.Q)
          THEN
            GVL_MSG_XTS.TransportMessageCtrl.Cmd    := E_MESSAGE_CTRL.MSG_CTRL_WRITE;
          END_IF
        END_IF
    END_CASE

  E_MESSAGE_STATE.MSG_STATE_WRITE:
    CASE eMsgProgress
    OF
      E_PROGRESS.PROGRESS_ERROR,
      E_PROGRESS.PROGRESS_DONE:
          tonIdleWriteMotion(IN := FALSE, PT:= tIdleWriteMotion);
        GVL_MSG_XTS.TransportMessageCtrl.Cmd        := E_MESSAGE_CTRL.MSG_CTRL_NULL;
    END_CASE

ELSE
    CASE eMsgProgress
    OF
      E_PROGRESS.PROGRESS_DONE:
          tonIdleWriteMotion(IN := FALSE, PT:= tIdleWriteMotion);
        GVL_MSG_XTS.TransportMessageCtrl.Cmd        := E_MESSAGE_CTRL.MSG_CTRL_NULL;
    END_CASE
END_CASE
//#################################################################################################################
// /application logging
//#################################################################################################################
GVL_MSG_XTS.ApplicationMessageData.Ctrl                         REF= GVL_MSG_XTS.ApplicationMessageCtrl;
GVL_MSG_XTS.ApplicationMessageData.State                        REF= GVL_MSG_XTS.ApplicationMessageState;

GVL_MSG_XTS.ApplicationMessageData.MessageIndex                 REF= GVL_MSG_XTS.MessageApplicationIndex;
GVL_MSG_XTS.ApplicationMessageData.ErrorIndex                   REF= GVL_MSG_XTS.MessageApplicationError;

GVL_MSG_XTS.ApplicationMessageData.DirRoot                      :=   ADR(GVL_MSG_XTS.LOG_DIR);
GVL_MSG_XTS.ApplicationMessageData.FileRoot                     :=   ADR(GVL_MSG_XTS.LOG_FILE_APP);
GVL_MSG_XTS.ApplicationMessageData.MsgList                      :=   ADR(GVL_MSG_XTS.ApplicationMessages);
GVL_MSG_XTS.ApplicationMessageData.LocalTime                    :=   ADR(GVL_MSG_XTS.dtLocalTime);

GVL_MSG_XTS.ApplicationMessageData();

eMsgState                                       := f_GetState   (GVL_MSG_XTS.ApplicationMessageState.State);
eMsgProgress                                    := f_GetProgress(GVL_MSG_XTS.ApplicationMessageState.State);


CASE eMsgState
OF
  E_MESSAGE_STATE.MSG_STATE_NULL:
    CASE eMsgProgress
    OF
      E_PROGRESS.PROGRESS_INVALID:
        IF (GVL_MSG_XTS.MessageApplicationIndex > GVL_MSG_XTS.MAX_MESSAGE/13) OR
           (GVL_MSG_XTS.MessageApplicationError > 0)
        THEN
          GVL_MSG_XTS.ApplicationMessageCtrl.Cmd                := E_MESSAGE_CTRL.MSG_CTRL_WRITE;
        ELSE
          tonIdleWriteApplication(IN := TRUE, PT:= tIdleWriteApplication);
          IF (tonIdleWriteApplication.Q)
          THEN
            GVL_MSG_XTS.ApplicationMessageCtrl.Cmd              := E_MESSAGE_CTRL.MSG_CTRL_WRITE;
          END_IF
        END_IF
    END_CASE

  E_MESSAGE_STATE.MSG_STATE_WRITE:
    CASE eMsgProgress
    OF
      E_PROGRESS.PROGRESS_ERROR,
      E_PROGRESS.PROGRESS_DONE:
        tonIdleWriteApplication(IN := FALSE, PT:= tIdleWriteApplication);
        GVL_MSG_XTS.ApplicationMessageCtrl.Cmd                  := E_MESSAGE_CTRL.MSG_CTRL_NULL;
    END_CASE

ELSE
    CASE eMsgProgress
    OF
      E_PROGRESS.PROGRESS_DONE:
        tonIdleWriteApplication(IN := FALSE, PT:= tIdleWriteApplication);
        GVL_MSG_XTS.ApplicationMessageCtrl.Cmd                  := E_MESSAGE_CTRL.MSG_CTRL_NULL;
    END_CASE
END_CASE
//#################################################################################################################
// logging/
//#################################################################################################################
//#################################################################################################################
//  /Transport Metrics
//#################################################################################################################
GVL_MSG_XTS.MetricsMessageData.Ctrl                             REF= GVL_MSG_XTS.MetricsMessageCtrl;
GVL_MSG_XTS.MetricsMessageData.State                            REF= GVL_MSG_XTS.MetricsMessageState;

GVL_MSG_XTS.MetricsMessageData.MessageIndex                     REF= GVL_MSG_XTS.MessageMetricsIndex;
GVL_MSG_XTS.MetricsMessageData.ErrorIndex                       REF= GVL_MSG_XTS.MessageMetricsError;

GVL_MSG_XTS.MetricsMessageData.DirRoot                          :=   ADR(GVL_MSG_XTS.LOG_DIR);
GVL_MSG_XTS.MetricsMessageData.FileRoot                         :=   ADR(GVL_MSG_XTS.LOG_FILE_METRIC);
GVL_MSG_XTS.MetricsMessageData.MsgList                          :=   ADR(GVL_MSG_XTS.MetricsMessages);
GVL_MSG_XTS.MetricsMessageData.LocalTime                        :=   ADR(GVL_MSG_XTS.dtLocalTime);

GVL_MSG_XTS.MetricsMessageData();

eMtrState                                   := f_GetState   (GVL_MSG_XTS.MetricsMessageState.State);
eMtrProgress                                := f_GetProgress(GVL_MSG_XTS.MetricsMessageState.State);

CASE eMtrState
OF
  E_MESSAGE_STATE.MSG_STATE_NULL:
    CASE eMtrProgress
    OF
      E_PROGRESS.PROGRESS_INVALID:
        IF (GVL_MSG_XTS.MessageMetricsIndex > GVL_MSG_XTS.MAX_MESSAGE/5) OR
           (GVL_MSG_XTS.MessageMetricsError > 0)
        THEN
          GVL_MSG_XTS.MetricsMessageCtrl.Cmd                    := E_MESSAGE_CTRL.MSG_CTRL_WRITE;
        ELSE
          tonIdleWriteMetric(IN := TRUE, PT:= tIdleWriteMetric);
          IF (tonIdleWriteMetric.Q)
          THEN
            GVL_MSG_XTS.MetricsMessageCtrl.Cmd                  := E_MESSAGE_CTRL.MSG_CTRL_WRITE;
          END_IF
        END_IF
    END_CASE

  E_MESSAGE_STATE.MSG_STATE_WRITE:
    CASE eMtrProgress
    OF
      E_PROGRESS.PROGRESS_ERROR,
      E_PROGRESS.PROGRESS_DONE:
        tonIdleWriteMetric(IN := FALSE, PT:= tIdleWriteMetric);
        GVL_MSG_XTS.MetricsMessageCtrl.Cmd                      := E_MESSAGE_CTRL.MSG_CTRL_NULL;
    END_CASE
ELSE
    CASE eMtrProgress
    OF
      E_PROGRESS.PROGRESS_DONE:
        tonIdleWriteMetric(IN := FALSE, PT:= tIdleWriteMetric);
        GVL_MSG_XTS.MetricsMessageCtrl.Cmd                      := E_MESSAGE_CTRL.MSG_CTRL_NULL;
    END_CASE
END_CASE
//#################################################################################################################
//  Transport Metrics/
//#################################################################################################################
//#################################################################################################################
//#################################################################################################################

ACTION Init:
CASE eInit
OF
  E_PROGRESS.PROGRESS_INVALID:          // startup procedure for your application
    eInit                               := E_PROGRESS.PROGRESS_INIT;

  E_PROGRESS.PROGRESS_INIT:
      nProcess                                        := 1;
      tProcess[nProcess]                              := T#750MS;

      GVL_APPLICATION.Simulation[nProcess].HandshakeRoute:= E_PROCESS_HANDSHAKE.E_SHAKE_DOUBLE;

      GVL_APPLICATION.Simulation[nProcess].StationFirst  := 1;
      GVL_APPLICATION.Simulation[nProcess].StationLast   := 16;

      GVL_APPLICATION.Simulation[nProcess].TargetFirst   := 20;
      GVL_APPLICATION.Simulation[nProcess].TargetLast    := 35;
      GVL_APPLICATION.Simulation[nProcess].TargetMask    := 2#0001; // mask for target station

      GVL_APPLICATION.Simulation[nProcess].CheckRangeLow :=   10.0;
      GVL_APPLICATION.Simulation[nProcess].CheckRangeHigh:= 1600.0;

      //---------------------------------------------------------

      // 2

      //---------------------------------------------------------
      nProcess                                        := 3;
      tProcess[nProcess]                              := T#2400MS;

      GVL_APPLICATION.Simulation[nProcess].HandshakeRoute:= E_PROCESS_HANDSHAKE.E_SHAKE_DOUBLE;

      GVL_APPLICATION.Simulation[nProcess].StationFirst  := 20;
      GVL_APPLICATION.Simulation[nProcess].StationLast   := 35;

      GVL_APPLICATION.Simulation[nProcess].TargetFirst   := 37;
      GVL_APPLICATION.Simulation[nProcess].TargetLast    := 37;
      GVL_APPLICATION.Simulation[nProcess].TargetMask    := 2#0001; // mask for target station

      GVL_APPLICATION.Simulation[nProcess].CheckRangeLow := 9000.0;
      GVL_APPLICATION.Simulation[nProcess].CheckRangeHigh:= 12100.0;

      //---------------------------------------------------------
      nProcess                                        := 4;
      tProcess[nProcess]                              := T#0MS;

      GVL_APPLICATION.Simulation[nProcess].HandshakeRoute:= E_PROCESS_HANDSHAKE.E_SHAKE_SEND;

      GVL_APPLICATION.Simulation[nProcess].StationFirst  := 37;
      GVL_APPLICATION.Simulation[nProcess].StationLast   := 37;

      GVL_APPLICATION.Simulation[nProcess].TargetFirst   := 38;
      GVL_APPLICATION.Simulation[nProcess].TargetLast    := 38;
      GVL_APPLICATION.Simulation[nProcess].TargetMask    := 2#0001; // mask for target station

      GVL_APPLICATION.Simulation[nProcess].CheckRangeLow := 12850.0;
      GVL_APPLICATION.Simulation[nProcess].CheckRangeHigh:= 13000.0;

      //---------------------------------------------------------
      nProcess                                        := 5;
      tProcess[nProcess]                              := T#0MS;

      GVL_APPLICATION.Simulation[nProcess].HandshakeRoute:= E_PROCESS_HANDSHAKE.E_SHAKE_SEND;

      GVL_APPLICATION.Simulation[nProcess].StationFirst  := 38;
      GVL_APPLICATION.Simulation[nProcess].StationLast   := 38;

      GVL_APPLICATION.Simulation[nProcess].TargetFirst   := 39;
      GVL_APPLICATION.Simulation[nProcess].TargetLast    := 39;
      GVL_APPLICATION.Simulation[nProcess].TargetMask    := 2#0001; // mask for target station

      GVL_APPLICATION.Simulation[nProcess].CheckRangeLow := 13900.0;
      GVL_APPLICATION.Simulation[nProcess].CheckRangeHigh:= 14100.0;

      //---------------------------------------------------------
      nProcess                                        := 6;
      tProcess[nProcess]                              := T#0MS;

      GVL_APPLICATION.Simulation[nProcess].HandshakeRoute:= E_PROCESS_HANDSHAKE.E_SHAKE_SEND;

      GVL_APPLICATION.Simulation[nProcess].StationFirst  := 39;
      GVL_APPLICATION.Simulation[nProcess].StationLast   := 39;

      GVL_APPLICATION.Simulation[nProcess].TargetFirst   := 41;
      GVL_APPLICATION.Simulation[nProcess].TargetLast    := 52;
      GVL_APPLICATION.Simulation[nProcess].TargetMask    := 2#0001; // mask for target station

      GVL_APPLICATION.Simulation[nProcess].CheckRangeLow := 14200.0;
      GVL_APPLICATION.Simulation[nProcess].CheckRangeHigh:= 14400.0;

      //---------------------------------------------------------
      nProcess                                        := 7;
      tProcess[nProcess]                              := T#3200MS;

      GVL_APPLICATION.Simulation[nProcess].HandshakeRoute:= E_PROCESS_HANDSHAKE.E_SHAKE_FAST;

      GVL_APPLICATION.Simulation[nProcess].StationFirst  := 41;
      GVL_APPLICATION.Simulation[nProcess].StationLast   := 52;

      GVL_APPLICATION.Simulation[nProcess].TargetFirst   := 57;
      GVL_APPLICATION.Simulation[nProcess].TargetLast    := 57;
      GVL_APPLICATION.Simulation[nProcess].TargetMask    := 2#0001; // mask for target station

      GVL_APPLICATION.Simulation[nProcess].CheckRangeLow := 14400.0;
      GVL_APPLICATION.Simulation[nProcess].CheckRangeHigh:= 17000.0;

      //---------------------------------------------------------
      nProcess                                        := 8;
      tProcess[nProcess]                              := T#0MS;

      GVL_APPLICATION.Simulation[nProcess].HandshakeRoute:= E_PROCESS_HANDSHAKE.E_SHAKE_SEND;

      GVL_APPLICATION.Simulation[nProcess].StationFirst  := 57;
      GVL_APPLICATION.Simulation[nProcess].StationLast   := 57;

      GVL_APPLICATION.Simulation[nProcess].TargetFirst   := 58;
      GVL_APPLICATION.Simulation[nProcess].TargetLast    := 65;
      GVL_APPLICATION.Simulation[nProcess].TargetMask    := 2#0001; // mask for target station

      GVL_APPLICATION.Simulation[nProcess].CheckRangeLow := 17500.0;
      GVL_APPLICATION.Simulation[nProcess].CheckRangeHigh:= 18100.0;

      //---------------------------------------------------------
      nProcess                                        := 9;
      tProcess[nProcess]                              := T#3200MS;

      GVL_APPLICATION.Simulation[nProcess].HandshakeRoute:= E_PROCESS_HANDSHAKE.E_SHAKE_SINGLE;

      GVL_APPLICATION.Simulation[nProcess].StationFirst  := 58;
      GVL_APPLICATION.Simulation[nProcess].StationLast   := 65;

      GVL_APPLICATION.Simulation[nProcess].TargetFirst   := 70;
      GVL_APPLICATION.Simulation[nProcess].TargetLast    := 70;
      GVL_APPLICATION.Simulation[nProcess].TargetMask    := 2#0001; // mask for target station

      GVL_APPLICATION.Simulation[nProcess].CheckRangeLow := 19400.0;
      GVL_APPLICATION.Simulation[nProcess].CheckRangeHigh:= 20500.0;

      //---------------------------------------------------------
      nProcess                                        := 10;
      tProcess[nProcess]                              := T#0MS;

      GVL_APPLICATION.Simulation[nProcess].HandshakeRoute:= E_PROCESS_HANDSHAKE.E_SHAKE_SEND;

      GVL_APPLICATION.Simulation[nProcess].StationFirst  := 70;
      GVL_APPLICATION.Simulation[nProcess].StationLast   := 70;

      GVL_APPLICATION.Simulation[nProcess].TargetFirst   := 71;
      GVL_APPLICATION.Simulation[nProcess].TargetLast    := 82;
      GVL_APPLICATION.Simulation[nProcess].TargetMask    := 2#0001; // mask for target station

      GVL_APPLICATION.Simulation[nProcess].CheckRangeLow := 20600.0;
      GVL_APPLICATION.Simulation[nProcess].CheckRangeHigh:= 21400.0;

      //---------------------------------------------------------
      nProcess                                        := 12;
      tProcess[nProcess]                              := T#4600MS;

      GVL_APPLICATION.Simulation[nProcess].HandshakeRoute:= E_PROCESS_HANDSHAKE.E_SHAKE_DOUBLE;

      GVL_APPLICATION.Simulation[nProcess].StationFirst  := 71;
      GVL_APPLICATION.Simulation[nProcess].StationLast   := 82;

      GVL_APPLICATION.Simulation[nProcess].TargetFirst   := 91;
      GVL_APPLICATION.Simulation[nProcess].TargetLast    := 91;
      GVL_APPLICATION.Simulation[nProcess].TargetMask    := 2#0001; // mask for target station

      GVL_APPLICATION.Simulation[nProcess].CheckRangeLow := 21400.0;
      GVL_APPLICATION.Simulation[nProcess].CheckRangeHigh:= 22800.0;

      //---------------------------------------------------------
      nProcess                                        := 13;
      tProcess[nProcess]                              := T#00MS;

      GVL_APPLICATION.Simulation[nProcess].HandshakeRoute:= E_PROCESS_HANDSHAKE.E_SHAKE_SEND;

      GVL_APPLICATION.Simulation[nProcess].StationFirst  := 91;
      GVL_APPLICATION.Simulation[nProcess].StationLast   := 91;

      GVL_APPLICATION.Simulation[nProcess].TargetFirst   := 95;
      GVL_APPLICATION.Simulation[nProcess].TargetLast    := 95;
      GVL_APPLICATION.Simulation[nProcess].TargetMask    := 2#0001; // mask for target station

      GVL_APPLICATION.Simulation[nProcess].CheckRangeLow := 22800.0;
      GVL_APPLICATION.Simulation[nProcess].CheckRangeHigh:= 23500.0;

      //---------------------------------------------------------
      nProcess                                        := 14;
      tProcess[nProcess]                              := T#0MS;

      GVL_APPLICATION.Simulation[nProcess].HandshakeRoute:= E_PROCESS_HANDSHAKE.E_SHAKE_SEND;

      GVL_APPLICATION.Simulation[nProcess].StationFirst  := 95;
      GVL_APPLICATION.Simulation[nProcess].StationLast   := 95;

      GVL_APPLICATION.Simulation[nProcess].TargetFirst   := 120;
      GVL_APPLICATION.Simulation[nProcess].TargetLast    := 133;
      GVL_APPLICATION.Simulation[nProcess].TargetMask    := 2#0001; // mask for target station

      GVL_APPLICATION.Simulation[nProcess].CheckRangeLow := 24000.0;
      GVL_APPLICATION.Simulation[nProcess].CheckRangeHigh:= 24100.0;

      //---------------------------------------------------------
      nProcess                                        := 15;
      tProcess[nProcess]                              := T#2500MS;

      GVL_APPLICATION.Simulation[nProcess].HandshakeRoute:= E_PROCESS_HANDSHAKE.E_SHAKE_DOUBLE;

      GVL_APPLICATION.Simulation[nProcess].StationFirst  := 120;
      GVL_APPLICATION.Simulation[nProcess].StationLast   := 133;

      GVL_APPLICATION.Simulation[nProcess].TargetFirst   := 140;
      GVL_APPLICATION.Simulation[nProcess].TargetLast    := 140;
      GVL_APPLICATION.Simulation[nProcess].TargetMask    := 2#0001; // mask for target station

      GVL_APPLICATION.Simulation[nProcess].CheckRangeLow := 24200.0;
      GVL_APPLICATION.Simulation[nProcess].CheckRangeHigh:= 27500.0;

      //---------------------------------------------------------
      nProcess                                        := 16;
      tProcess[nProcess]                              := T#0MS;

      GVL_APPLICATION.Simulation[nProcess].HandshakeRoute:= E_PROCESS_HANDSHAKE.E_SHAKE_SEND;

      GVL_APPLICATION.Simulation[nProcess].StationFirst  := 140;
      GVL_APPLICATION.Simulation[nProcess].StationLast   := 140;

      GVL_APPLICATION.Simulation[nProcess].TargetFirst   := 141;
      GVL_APPLICATION.Simulation[nProcess].TargetLast    := 141;
      GVL_APPLICATION.Simulation[nProcess].TargetMask    := 2#0001; // mask for target station

      GVL_APPLICATION.Simulation[nProcess].CheckRangeLow := 27970.0;
      GVL_APPLICATION.Simulation[nProcess].CheckRangeHigh:= 1250.0;

      //---------------------------------------------------------
      nProcess                                        := 17;
      tProcess[nProcess]                              := T#0MS;

      GVL_APPLICATION.Simulation[nProcess].HandshakeRoute:= E_PROCESS_HANDSHAKE.E_SHAKE_SEND;

      GVL_APPLICATION.Simulation[nProcess].StationFirst  := 141;
      GVL_APPLICATION.Simulation[nProcess].StationLast   := 141;

      GVL_APPLICATION.Simulation[nProcess].TargetFirst   := 142;
      GVL_APPLICATION.Simulation[nProcess].TargetLast    := 142;
      GVL_APPLICATION.Simulation[nProcess].TargetMask    := 2#0001; // mask for target station

      GVL_APPLICATION.Simulation[nProcess].CheckRangeLow := 3950.0;
      GVL_APPLICATION.Simulation[nProcess].CheckRangeHigh:= 4100.0;

      //---------------------------------------------------------
      nProcess                                        := 18;
      tProcess[nProcess]                              := T#0MS;

      GVL_APPLICATION.Simulation[nProcess].HandshakeRoute:= E_PROCESS_HANDSHAKE.E_SHAKE_SEND;

      GVL_APPLICATION.Simulation[nProcess].StationFirst  := 142;
      GVL_APPLICATION.Simulation[nProcess].StationLast   := 142;

      GVL_APPLICATION.Simulation[nProcess].TargetFirst   := 20;
      GVL_APPLICATION.Simulation[nProcess].TargetLast    := 35;
      GVL_APPLICATION.Simulation[nProcess].TargetMask    := 2#0001; // mask for target station

      GVL_APPLICATION.Simulation[nProcess].CheckRangeLow := 4500.0;
      GVL_APPLICATION.Simulation[nProcess].CheckRangeHigh:= 5600.0;


    eInit                                                 := E_PROGRESS.PROGRESS_BUSY;

  E_PROGRESS.PROGRESS_BUSY:
    GVL_MSG_XTS.TransportMessageCtrl.Cmd                  := E_MESSAGE_CTRL.MSG_CTRL_INIT;
    GVL_MSG_XTS.MetricsMessageCtrl.Cmd                    := E_MESSAGE_CTRL.MSG_CTRL_INIT;
    eInit                                                 := E_PROGRESS.PROGRESS_PREPARE;

  E_PROGRESS.PROGRESS_PREPARE:
    eInit                                                 := E_PROGRESS.PROGRESS_STARTUP;

  E_PROGRESS.PROGRESS_STARTUP:
    eInit                                                 := E_PROGRESS.PROGRESS_DONE;
    FOR nProcess := 1 TO MAX_PROCESS
    DO
      IF (GVL_APPLICATION.Simulation[nProcess].StationCount > 0)
      THEN
        GVL_APPLICATION.Simulation[nProcess].EnableProcess := TO_DWORD(EXPT(2,GVL_APPLICATION.Simulation[nProcess].StationCount))-1;
        GVL_APPLICATION.Simulation[nProcess].MoverEnter    := TRUE;
        GVL_APPLICATION.Simulation[nProcess].MoverOut      := TRUE;

      END_IF
    END_FOR
END_CASE
END_ACTION

END_PROGRAM

// ---- _types/f_GetState.TcPOU
// global function to extract state identifier from combined value
FUNCTION f_GetState : uint
VAR_INPUT
  state     : UINT; // combined value of identifier + e_progress
END_VAR
VAR
  _stx      : uint;
END_VAR

_stx          := state MOD E_PROGRESS.PROGRESS_INIT;

IF (_stx = 0)
THEN
  f_GetState  := state;
ELSE
  f_GetState  := _stx;
END_IF

END_FUNCTION

// ---- _types/f_GetProgress.TcPOU
// global function to extract e_progress from combined value
FUNCTION f_GetProgress : uint
VAR_INPUT
  state     : UINT;
END_VAR
VAR
  nP        : uint;
END_VAR


nP := state / E_PROGRESS.PROGRESS_INIT;

f_GetProgress := nP * E_PROGRESS.PROGRESS_INIT;

END_FUNCTION

// ---- MAPPING/MAPPING_XTS_out.TcPOU
PROGRAM MAPPING_XTS_out
VAR
  sMapping              : STRING;
  bFirstCycle           : BOOL := TRUE;

  YardState             : U_YARD_STATE;
  InstanceState         : U_INSTANCE_STATE;
  TicketListOutput      : U_TICKET_LIST_DATA_OUTPUT;
  TicketListState       : U_TICKET_LIST_STATE;

  TransportControl      : U_XTS_TRANSPORT_CTRL;
  StationControl        : U_XTS_STATION_CTRL;


  szTransportCtrl       : ARRAY[1..2] OF UDINT;
  szStationControl      : ARRAY[1..2] OF UDINT;
END_VAR


IF (bFirstCycle)
THEN
  bFirstCycle             := FALSE;

  szTransportCtrl[1]      := SIZEOF(TransportControl);
  szTransportCtrl[2]      := SIZEOF(GVL_XTS.XtsTransportCtrl);

  szStationControl[1]     := SIZEOF(StationControl);
  szStationControl[2]     := SIZEOF(GVL_XTS.StationCtrl);
END_IF
//---------------------------------------------------------------------
IF (SIZEOF(TransportControl) <> SIZEOF(GVL_XTS.XtsTransportCtrl))
THEN
  sMapping  := 'TransportControl sizes DO NOT match';
  RETURN;
END_IF
//---------------------------------------------------------------------
IF (SIZEOF(StationControl) <> SIZEOF(GVL_XTS.StationCtrl))
THEN
  sMapping  := 'StationControl sizes DO NOT match';
  RETURN;
END_IF
//---------------------------------------------------------------------
IF (SIZEOF(YardState) <> SIZEOF(GVL_APPLICATION.YardState))
THEN
  sMapping  := 'YardState sizes DO NOT match';
  RETURN;
END_IF
//---------------------------------------------------------------------
IF (SIZEOF(InstanceState) <> SIZEOF(GVL_APPLICATION.InstanceState))
THEN
  sMapping  := 'InstanceState sizes DO NOT match';
  RETURN;
END_IF
//---------------------------------------------------------------------
sMapping    := 'MAPPING_XTS_OUTPUT ACTIVE';
//-----------------------------------------------------------------------------------------------------
//       destination,           source,                             size
//-----------------------------------------------------------------------------------------------------
  memcpy(ADR(TransportControl), ADR(GVL_XTS.XtsTransportCtrl),      SIZEOF(TransportControl));
  memcpy(ADR(StationControl),   ADR(GVL_XTS.StationCtrl),           SIZEOF(StationControl));
//-----------------------------------------------------------------------------------------------------
//-----------------------------------------------------------------------------------------------------
//       destination,           source,                                     size
//-----------------------------------------------------------------------------------------------------
  memcpy(ADR(YardState),        ADR(GVL_APPLICATION.YardState),             SIZEOF(YardState));
  memcpy(ADR(InstanceState),    ADR(GVL_APPLICATION.InstanceState),         SIZEOF(InstanceState));
  memcpy(ADR(TicketListState),  ADR(GVL_APPLICATION.TicketListState),       SIZEOF(TicketListState));
  memcpy(ADR(TicketListOutput), ADR(GVL_APPLICATION.TicketListDataOutput),  SIZEOF(TicketListOutput));
//-----------------------------------------------------------------------------------------------------
//-----------------------------------------------------------------------------------------------------

END_PROGRAM

// ---- APPLICATION/_types/YardMaster/fb_YardMaster.TcPOU
//---------------------------------------------------------------------------------------------------------------
//
//  HAUD 2025.11.03
//
//  fb_YardMaster
// 
//  - top level organizer for the transport system
//
//  - commands TransportUnit
//    - subsumes commands into sequences
//    - reports to higher up (TowerControl)
//
//  - initializes Collectors
//    - Collectors initialize their range of stations
// 
//---------------------------------------------------------------------------------------------------------------
FUNCTION_BLOCK fb_YardMaster
VAR
  _eCheck                       : E_YARD_CHECK;
  _eInit                        : E_PROGRESS;

  _Ctrl                         : REFERENCE TO ST_YARD_CTRL;
  _State                        : REFERENCE TO ST_YARD_STATE;

  _eResult                      : E_PROGRESS;

  _eCmd,
  _eCmdOld                      : E_INSTANCE_CMD;
  _eState                       : E_INSTANCE_STATE;

  // Transport Ctrl/State
  _XtsTransportCtrl             : REFERENCE TO ST_XTS_TRANSPORT_CTRL;
  _XtsTransportState            : REFERENCE TO ST_XTS_TRANSPORT_STATE;

  _ItfCollectors                : ARRAY[1..MAX_PROCESS] OF I_ProcessCollector;

  _ItfTicketList                : I_Process_LinkedList;

  _stMsg                        : ST_Message;
  _MessageLevel                 : E_MessageType := E_MessageType.eMessageInfo;
END_VAR

IF NOT Check() THEN RETURN; END_IF
//-----------------------------------------------------------------------------
//-----------------------------------------------------------------------------
// set message device
//-----------------------------------------------------------------------------
_stMsg.eDevice                  := e_Device.YardMaster;
//-----------------------------------------------------------------------------
_eCmd                           := _Ctrl.Cmd;
// check for command change
// get state for cmd
IF (_eCmd <> _eCmdOld)
THEN
  _eState                       := Cmd(_eCmd);
  _eCmdOld                      := _eCmd;

  IF (_MessageLevel > E_MessageType.eMessageError)
  THEN
    _stMsg.eType                := E_MessageType.eMessageInfo;
    _stMsg.eSubdevice           := e_Subdevice.Application_Cmd;
    _stMsg.iErrorNumber         := 0;
    _stMsg.sText                := concat(TO_STRING(_eCmd), ': ');
    _stMsg.sText                := concat(_stMsg.sText,  TO_STRING(_eState));
    f_MessageSet(_stMsg);
  END_IF

END_IF

CASE _eResult
OF
  E_PROGRESS.PROGRESS_INVALID:
    _State.State                := TO_UINT(_eResult);

  E_PROGRESS.PROGRESS_ERROR:
    _State.State                := _eState + E_PROGRESS.PROGRESS_ERROR;

  E_PROGRESS.PROGRESS_DONE:
    _State.State                := _eState + E_PROGRESS.PROGRESS_DONE;

ELSE
  _State.State                  := _eState + _eResult;

  CASE _eState
  OF
    E_INSTANCE_STATE.INIT:
      _eInit := _eResult        := Init(TRUE);

    E_INSTANCE_STATE.DISABLED:
      _eResult                  := Disable(TRUE);
  
    E_INSTANCE_STATE.ENABLED:
      _eResult                  := Enable(TRUE);

    E_INSTANCE_STATE.CLEARED:
      _eResult                  := Clear(TRUE);

    E_INSTANCE_STATE.WORKING:
      _eResult                  := Work(TRUE);

  ELSE
    _eResult                    := E_PROGRESS.PROGRESS_INVALID;
  END_CASE
END_CASE
//-----------------------------------------------------------------------------
//-----------------------------------------------------------------------------
_State.TransportState           := _XtsTransportState;
//-----------------------------------------------------------------------------
//-----------------------------------------------------------------------------

METHOD Check : BOOL
VAR_INST
  _nIdx       : E_INSTANCE;
END_VAR
//-----------------------------------------------------------------------------
//-----------------------------------------------------------------------------
// reference checks
//-----------------------------------------------------------------------------
IF NOT __ISVALIDREF(_Ctrl)
THEN
  _eCheck                   := E_YARD_CHECK.POINTER_CTRL_INVALID;
  RETURN;
END_IF

IF NOT __ISVALIDREF(_State)
THEN
  _eCheck                   := E_YARD_CHECK.POINTER_STATE_INVALID;
  RETURN;
END_IF

IF NOT __ISVALIDREF(_XtsTransportCtrl)
THEN
  _eCheck                   := E_YARD_CHECK.POINTER_TRANSPORT_CTRL_INVALID;
  RETURN;
END_IF

IF NOT __ISVALIDREF(_XtsTransportState)
THEN
  _eCheck                   := E_YARD_CHECK.POINTER_TRANSPORT_STATE_INVALID;
  RETURN;
END_IF

FOR _nIdx := 1 TO MAX_PROCESS
DO
  IF NOT (_ItfCollectors[_nIdx] <> 0)
  THEN
    _eCheck                 := E_YARD_CHECK.POINTER_COLLECTOR_ITF_INVALID;
    RETURN;
  END_IF
END_FOR

IF NOT (_ItfTicketList <> 0)
THEN
  _eCheck                   := E_YARD_CHECK.REFERENCE_TICKET_LIST_ITF_INVALID;
  RETURN;
END_IF

//-----------------------------------------------------------------------------
//-----------------------------------------------------------------------------
_eCheck                     := E_YARD_CHECK.CHECK_DONE;
Check                       := TRUE;
END_METHOD

METHOD Clear : E_PROGRESS
VAR_INPUT
  Execute     : BOOL;
END_VAR
VAR_INST
  _nErrorId   : UDINT;
  _eResult,
  _eState     : E_PROGRESS;

  _nIdx       : UINT;
  _eInstance  : E_INSTANCE;
END_VAR
//-----------------------------------------------------------------------------
IF NOT Execute 
THEN 
	_eState                       := E_PROGRESS.PROGRESS_INIT; 
END_IF 
//-----------------------------------------------------------------------------
IF NOT Check() 
THEN 
	Clear                         := E_PROGRESS.PROGRESS_ERROR; 
	RETURN; 
END_IF
//-----------------------------------------------------------------------------
//-----------------------------------------------------------------------------
CASE _eState
OF
  //---------------------------------------------------------------------------------------------------------------
  //---------------------------------------------------------------------------------------------------------------
  E_PROGRESS.PROGRESS_INIT:     // startup procedure for your application
    IF Execute
    THEN
      _nIdx                     := 1;
      _eState                   := E_PROGRESS.PROGRESS_BUSY;
  
      IF (_MessageLevel > E_MessageType.eMessageError)
      THEN
        _stMsg.eType            := E_MessageType.eMessageInfo;
        _stMsg.eSubdevice       := e_Subdevice.Application_Clear;
        _stMsg.iErrorNumber     := 0;
        _stMsg.sText            := concat(TO_STRING(_eState), ': ');
        f_MessageSet(_stMsg);
      END_IF
    END_IF

  //---------------------------------------------------------------------------------------------------------------
  //---------------------------------------------------------------------------------------------------------------
  E_PROGRESS.PROGRESS_BUSY:
    _XtsTransportCtrl.Cmd                 := E_XTS_TRANSPORT_CTRL.CMD_GROUP_CLEAR;

    IF (_XtsTransportState.State > E_PROGRESS.PROGRESS_ERROR)
    THEN
      _eState                             := E_PROGRESS.PROGRESS_PREPARE;
    END_IF
  //---------------------------------------------------------------------------------------------------------------
  //---------------------------------------------------------------------------------------------------------------
  E_PROGRESS.PROGRESS_PREPARE:
    _XtsTransportCtrl.Cmd                 := E_XTS_TRANSPORT_CTRL.CMD_MOVER_STOP;

    IF (_XtsTransportState.State > E_PROGRESS.PROGRESS_ERROR)
    THEN
      _eState                             := E_PROGRESS.PROGRESS_STARTUP;
    END_IF
  //---------------------------------------------------------------------------------------------------------------
  //---------------------------------------------------------------------------------------------------------------
  E_PROGRESS.PROGRESS_STARTUP:
    _XtsTransportCtrl.Cmd                 := E_XTS_TRANSPORT_CTRL.CMD_GROUP_CLEAR;

    IF (_XtsTransportState.State = E_XTS_TRANSPORT_STATE.TRANSPORT_GROUP_CLEAR + E_PROGRESS.PROGRESS_ERROR)
    THEN
      _eState                             := E_PROGRESS.PROGRESS_PREPARE;

    ELSIF (_XtsTransportState.State = E_XTS_TRANSPORT_STATE.TRANSPORT_GROUP_CLEAR + E_PROGRESS.PROGRESS_DONE)
    THEN 
      _eState                             := E_PROGRESS.PROGRESS_CHECK;
    END_IF
  //---------------------------------------------------------------------------------------------------------------
  //---------------------------------------------------------------------------------------------------------------
  E_PROGRESS.PROGRESS_CHECK:
    _eResult                              := _ItfCollectors[_nIdx].Init(FALSE);
    _eState                               := E_PROGRESS.PROGRESS_OCCUPIED;
  //---------------------------------------------------------------------------------------------------------------
  //---------------------------------------------------------------------------------------------------------------
  E_PROGRESS.PROGRESS_OCCUPIED:
    _eResult                              := _ItfCollectors[_nIdx].Init(TRUE);

    IF (_eResult = E_PROGRESS.PROGRESS_DONE)
    THEN
      _eState                             := E_PROGRESS.PROGRESS_WORKING;
    END_IF
  //---------------------------------------------------------------------------------------------------------------
  //---------------------------------------------------------------------------------------------------------------
  E_PROGRESS.PROGRESS_WORKING:
    IF NOT (_nIdx < GVL_APPLICATION.MAX_PROCESS)
    THEN
      _eState                     := E_PROGRESS.PROGRESS_STILL_WORKING;
    ELSE
      _nIdx                       := _nIdx + 1;
      _eState                     := E_PROGRESS.PROGRESS_CHECK;
    END_IF
  //---------------------------------------------------------------------------------------------------------------
  //---------------------------------------------------------------------------------------------------------------
  E_PROGRESS.PROGRESS_STILL_WORKING:
    _eState                     := E_PROGRESS.PROGRESS_DONE;

    IF (_MessageLevel > E_MessageType.eMessageError)
    THEN
      _stMsg.eType              := E_MessageType.eMessageInfo;
      _stMsg.eSubdevice         := e_Subdevice.Application_Clear;
      _stMsg.iErrorNumber       := 0;
      _stMsg.sText              := concat(TO_STRING(_eState), ': ');
      f_MessageSet(_stMsg);
    END_IF

END_CASE
//-----------------------------------------------------------------------------
//-----------------------------------------------------------------------------
Clear                           := _eState;
END_METHOD

METHOD PRIVATE Cmd : E_INSTANCE_STATE
VAR_INPUT
  Command   : E_INSTANCE_CMD;
END_VAR
VAR_INST
  _eRslt    : E_PROGRESS;
  _eState   : E_INSTANCE_STATE;
END_VAR
IF NOT Check() THEN RETURN; END_IF


CASE Command
OF
  E_INSTANCE_CMD.NULL:  // clear all method calls
    _eState                   := E_INSTANCE_STATE.NULL;
    _eRslt                    := Init    (FALSE);
    _eRslt                    := Disable (FALSE);
    _eRslt                    := Enable  (FALSE);
    _eRslt                    := Clear   (FALSE);

  E_INSTANCE_CMD.INIT:  // clear methods for initialization
    _eState                   := E_INSTANCE_STATE.INIT;
    _eResult                  := Init(FALSE);

ELSE
  IF NOT (_eInit = E_PROGRESS.PROGRESS_DONE)
  THEN
    // no init, no further commands possible
    _eState                   := E_INSTANCE_STATE.INVALID;

    _stMsg.eType              := E_MessageType.eMessageWarning;
    _stMsg.eSubdevice         := e_Subdevice.Application_Cmd;
    _stMsg.iErrorNumber       := Command;
    _stMsg.sText              := concat('_eInit: ', TO_STRING(_eInit));
    _stMsg.sText              := concat(_stMsg.sText, ': ');
    _stMsg.sText              := concat(_stMsg.sText, TO_STRING(_eState));
    f_MessageSet(_stMsg);

  ELSE
    CASE Command
    OF
      E_INSTANCE_CMD.DISABLE:
        _eState               := E_INSTANCE_STATE.DISABLED;
        _eResult              := Disable (FALSE);

      E_INSTANCE_CMD.ENABLE:
        _eState               := E_INSTANCE_STATE.ENABLED;
        _eResult              := Enable  (FALSE);

      E_INSTANCE_CMD.CLEAR:
        _eState               := E_INSTANCE_STATE.CLEARED;
        _eResult              := Clear   (FALSE);

      E_INSTANCE_CMD.WORK:
        _eState               := E_INSTANCE_STATE.WORKING;
        _eResult              := Work    (FALSE);

    ELSE
        _eState               := E_INSTANCE_STATE.INVALID;

        _stMsg.eType          := E_MessageType.eMessageError;
        _stMsg.eSubdevice     := e_Subdevice.Application_Cmd;
        _stMsg.iErrorNumber   := Command;
        _stMsg.sText          := concat('Command: ', TO_STRING(Command));
        _stMsg.sText          := concat(_stMsg.sText, ': ');
        _stMsg.sText          := concat(_stMsg.sText, TO_STRING(_eState));
        f_MessageSet(_stMsg);
    END_CASE
  END_IF
END_CASE

Cmd                           := _eState;
END_METHOD

PROPERTY CollectorInterfaces : array[1..MAX_PROCESS] of I_ProcessCollector
SET
_ItfCollectors := CollectorInterfaces;
END_SET
END_PROPERTY

PROPERTY Ctrl : REFERENCE TO ST_YARD_CTRL
SET
_Ctrl REF= Ctrl;
END_SET
END_PROPERTY

METHOD Disable : E_PROGRESS // RemoveAllAxis from CA Group, disable CA Group, disable all movers
VAR_INPUT
  Execute     : BOOL;
END_VAR
VAR_INST
  _nErrorId   : UDINT;
  _eState     : E_PROGRESS;
END_VAR
//-----------------------------------------------------------------------------
IF NOT Execute 
THEN 
	_eState                       := E_PROGRESS.PROGRESS_INIT; 
END_IF 
//-------------------------------------------------------------------------------
IF NOT Check() 
THEN 
	Disable                       := E_PROGRESS.PROGRESS_ERROR; 
	RETURN; 
END_IF
//-------------------------------------------------------------------------------
//-------------------------------------------------------------------------------
CASE _eState
OF
  E_PROGRESS.PROGRESS_INIT:
    IF Execute
    THEN
      _nErrorId                 := 0;

      _XtsTransportCtrl.Cmd     := E_XTS_TRANSPORT_CTRL.CMD_NULL;
      _eState                   := E_PROGRESS.PROGRESS_BUSY;

      IF (_MessageLevel > E_MessageType.eMessageError)
      THEN
        _stMsg.eType            := E_MessageType.eMessageInfo;
        _stMsg.eSubdevice       := e_Subdevice.Application_Disable;
        _stMsg.iErrorNumber     := 0;
        _stMsg.sText            := concat(TO_STRING(_eState), ': ');
        f_MessageSet(_stMsg);
      END_IF
    END_IF
  //-----------------------------------------------------------------------------
  //-----------------------------------------------------------------------------
  E_PROGRESS.PROGRESS_BUSY:
    _XtsTransportCtrl.Cmd       := E_XTS_TRANSPORT_CTRL.CMD_GROUP_CLEAR; 
    _eState                     := E_PROGRESS.PROGRESS_PREPARE;
  //-----------------------------------------------------------------------------
  //-----------------------------------------------------------------------------
  E_PROGRESS.PROGRESS_PREPARE:
    IF (_XtsTransportState.State = E_XTS_TRANSPORT_STATE.TRANSPORT_GROUP_CLEAR + E_PROGRESS.PROGRESS_ERROR)
    THEN
      _eState                   := E_PROGRESS.PROGRESS_BUSY;
      _XtsTransportCtrl.Cmd     := E_XTS_TRANSPORT_CTRL.CMD_NULL;

      _nErrorId                 := _XtsTransportState.GroupInfo.GroupErrorId; 

    ELSIF (_XtsTransportState.State = E_XTS_TRANSPORT_STATE.TRANSPORT_GROUP_CLEAR + E_PROGRESS.PROGRESS_DONE)
    THEN
      _eState                   := E_PROGRESS.PROGRESS_STARTUP;
    END_IF
  //-----------------------------------------------------------------------------
  //-----------------------------------------------------------------------------
  E_PROGRESS.PROGRESS_STARTUP:
    _XtsTransportCtrl.Cmd       := E_XTS_TRANSPORT_CTRL.CMD_MOVER_DISABLE; 
    _eState                     := E_PROGRESS.PROGRESS_CHECK;
  //-----------------------------------------------------------------------------
  //-----------------------------------------------------------------------------
  E_PROGRESS.PROGRESS_CHECK:
    IF (_XtsTransportState.State = E_XTS_TRANSPORT_STATE.TRANSPORT_MOVER_DISABLE + E_PROGRESS.PROGRESS_ERROR)
    THEN
      _eState                   := E_PROGRESS.PROGRESS_ERROR;

      _stMsg.eType              := E_MessageType.eMessageError;
      _stMsg.eSubdevice         := e_Subdevice.Application_Disable;
      _stMsg.iErrorNumber       := 0;
      _stMsg.sText              := concat(TO_STRING(_eState), ': ');
      f_MessageSet(_stMsg);

    ELSIF (_XtsTransportState.State = E_XTS_TRANSPORT_STATE.TRANSPORT_MOVER_DISABLE + E_PROGRESS.PROGRESS_DONE)
    THEN
      _eState                   := E_PROGRESS.PROGRESS_DONE;

      IF (_MessageLevel > E_MessageType.eMessageError)
      THEN
        _stMsg.eType            := E_MessageType.eMessageInfo;
        _stMsg.eSubdevice       := e_Subdevice.Application_Disable;
        _stMsg.iErrorNumber     := 0;
        _stMsg.sText            := concat(TO_STRING(_eState), ': ');
        f_MessageSet(_stMsg);
      END_IF
    END_IF
END_CASE
//-------------------------------------------------------------------------------
//-------------------------------------------------------------------------------

Disable                         := _eState;
END_METHOD

METHOD Enable : E_PROGRESS // AddAllAxis to CA Group, Enable CA Group, Enable all movers
VAR_INPUT
  Execute     : BOOL;
END_VAR
VAR_INST
  _nErrorId   : UDINT;
  _eState     : E_PROGRESS;
END_VAR
//-----------------------------------------------------------------------------
IF NOT Execute 
THEN 
	_eState                       := E_PROGRESS.PROGRESS_INIT; 
END_IF 
//-----------------------------------------------------------------------------
IF NOT Check() 
THEN 
	Enable                        := E_PROGRESS.PROGRESS_ERROR; 
	RETURN; 
END_IF
//-----------------------------------------------------------------------------
//-----------------------------------------------------------------------------
CASE _eState
OF
  E_PROGRESS.PROGRESS_INIT:
    IF Execute
    THEN
      _nErrorId                 := 0;

      _XtsTransportCtrl.Cmd     := E_XTS_TRANSPORT_CTRL.CMD_NULL;
      _eState                   := E_PROGRESS.PROGRESS_BUSY;

      IF (_MessageLevel > E_MessageType.eMessageError)
      THEN
        _stMsg.eType            := E_MessageType.eMessageInfo;
        _stMsg.eSubdevice       := e_Subdevice.Application_Enable;
        _stMsg.iErrorNumber     := 0;
        _stMsg.sText            := concat(TO_STRING(_eState), ': ');
        f_MessageSet(_stMsg);
      END_IF
    END_IF
  //-----------------------------------------------------------------------------
  //-----------------------------------------------------------------------------
  E_PROGRESS.PROGRESS_BUSY:
    _XtsTransportCtrl.Cmd       := E_XTS_TRANSPORT_CTRL.CMD_GROUP_CLEAR;

    IF (_XtsTransportState.State = E_XTS_TRANSPORT_STATE.TRANSPORT_GROUP_CLEAR + E_PROGRESS.PROGRESS_ERROR)
    THEN
      _eState                   := E_PROGRESS.PROGRESS_ERROR;
      _nErrorId                 := _XtsTransportState.GroupInfo.GroupErrorId; 

    ELSIF (_XtsTransportState.State = E_XTS_TRANSPORT_STATE.TRANSPORT_GROUP_CLEAR + E_PROGRESS.PROGRESS_DONE)
    THEN
      _eState                   := E_PROGRESS.PROGRESS_PREPARE;
    END_IF
  //-----------------------------------------------------------------------------
  //-----------------------------------------------------------------------------
  E_PROGRESS.PROGRESS_PREPARE:
    _XtsTransportCtrl.Cmd       := E_XTS_TRANSPORT_CTRL.CMD_GROUP_BUILD;

    IF (_XtsTransportState.State = E_XTS_TRANSPORT_STATE.TRANSPORT_GROUP_BUILD + E_PROGRESS.PROGRESS_ERROR)
    THEN
      _eState                   := E_PROGRESS.PROGRESS_ERROR;
      _nErrorId                 := _XtsTransportState.GroupInfo.GroupErrorId; 

    ELSIF (_XtsTransportState.State = E_XTS_TRANSPORT_STATE.TRANSPORT_GROUP_BUILD + E_PROGRESS.PROGRESS_DONE)
    THEN
      _eState                   := E_PROGRESS.PROGRESS_STARTUP;
    END_IF
  //-----------------------------------------------------------------------------
  //-----------------------------------------------------------------------------
  E_PROGRESS.PROGRESS_STARTUP:
    _XtsTransportCtrl.Cmd       := E_XTS_TRANSPORT_CTRL.CMD_MOVER_ENABLE; 
    _eState                     := E_PROGRESS.PROGRESS_CHECK;
  //-----------------------------------------------------------------------------
  //-----------------------------------------------------------------------------
  E_PROGRESS.PROGRESS_CHECK:
    IF (_XtsTransportState.State = E_XTS_TRANSPORT_STATE.TRANSPORT_MOVER_ENABLE + E_PROGRESS.PROGRESS_ERROR)
    THEN
      _eState                   := E_PROGRESS.PROGRESS_ERROR;

    ELSIF (_XtsTransportState.State = E_XTS_TRANSPORT_STATE.TRANSPORT_MOVER_ENABLE + E_PROGRESS.PROGRESS_DONE)
    THEN
      _eState                   := E_PROGRESS.PROGRESS_OCCUPIED;
    END_IF
  //-----------------------------------------------------------------------------
  //-----------------------------------------------------------------------------
  E_PROGRESS.PROGRESS_OCCUPIED:
    _XtsTransportCtrl.Cmd       := E_XTS_TRANSPORT_CTRL.CMD_GROUP_ENABLE; 
    _eState                     := E_PROGRESS.PROGRESS_WORKING;
  //-----------------------------------------------------------------------------
  //-----------------------------------------------------------------------------
  E_PROGRESS.PROGRESS_WORKING:
    IF (_XtsTransportState.State = E_XTS_TRANSPORT_STATE.TRANSPORT_GROUP_ENABLE + E_PROGRESS.PROGRESS_ERROR)
    THEN
      _eState                   := E_PROGRESS.PROGRESS_ERROR;

      _stMsg.eType              := E_MessageType.eMessageError;
      _stMsg.eSubdevice         := e_Subdevice.Application_Enable;
      _stMsg.iErrorNumber       := 0;
      _stMsg.sText              := concat(TO_STRING(_eState), ': ');
      f_MessageSet(_stMsg);

    ELSIF (_XtsTransportState.State = E_XTS_TRANSPORT_STATE.TRANSPORT_GROUP_ENABLE + E_PROGRESS.PROGRESS_DONE)
    THEN
      _eState                   := E_PROGRESS.PROGRESS_DONE;

      IF (_MessageLevel > E_MessageType.eMessageError)
      THEN
        _stMsg.eType            := E_MessageType.eMessageInfo;
        _stMsg.eSubdevice       := e_Subdevice.Application_Enable;
        _stMsg.iErrorNumber     := 0;
        _stMsg.sText            := concat(TO_STRING(_eState), ': ');
        f_MessageSet(_stMsg);
      END_IF
    END_IF
END_CASE
//-----------------------------------------------------------------------------
//-----------------------------------------------------------------------------

Enable                          := _eState;
END_METHOD

METHOD Init       : E_PROGRESS  
VAR_INPUT
  Execute         : BOOL;
END_VAR
VAR_INST
  _nInstance      : UINT;
  _nInstanceError : E_INSTANCE;
  _nIdx,
  _nErrorId       : UDINT;
  _eResult        : E_PROGRESS;
  _eState         : E_PROGRESS;
END_VAR
//------------------------------------------------------------------------------------------------------
IF NOT Execute 
THEN 
	_eState                                 := E_PROGRESS.PROGRESS_INIT; 
END_IF 
//------------------------------------------------------------------------------------------------------
IF NOT Check() 
THEN 
	Init                                    := E_PROGRESS.PROGRESS_ERROR; 
	RETURN; 
END_IF
//-------------------------------------------------------------------------------------------------------
//-------------------------------------------------------------------------------------------------------
CASE _eState
OF
  //-----------------------------------------------------------------------------------------------------
  //-----------------------------------------------------------------------------------------------------
  E_PROGRESS.PROGRESS_INIT:               // startup procedure for your application
    IF Execute
    THEN
      _nInstance                          := 1;
      _nInstanceError                     := E_INSTANCE.INSTANCE_NULL;
      _eState                             := E_PROGRESS.PROGRESS_BUSY;
      _XtsTransportCtrl.Cmd               := E_XTS_TRANSPORT_CTRL.CMD_NULL;

      IF (_MessageLevel > E_MessageType.eMessageError)
      THEN
        _stMsg.eType                      := E_MessageType.eMessageInfo;
        _stMsg.eSubdevice                 := e_Subdevice.Application_Init;
        _stMsg.iErrorNumber               := 0;
        _stMsg.sText                      := concat(TO_STRING(_eState), ': ');
        f_MessageSet(_stMsg);
      END_IF

      FOR _nIdx := 1 TO MAX_PROCESS
      DO
        _eResult                          := _ItfCollectors[_nIdx].Init(FALSE);
      END_FOR
    END_IF
  //-----------------------------------------------------------------------------------------------------
  //-----------------------------------------------------------------------------------------------------
  E_PROGRESS.PROGRESS_BUSY:
    _XtsTransportCtrl.Cmd                 := E_XTS_TRANSPORT_CTRL.CMD_INIT;
    IF (_XtsTransportState.State = E_XTS_TRANSPORT_STATE.TRANSPORT_INIT + E_PROGRESS.PROGRESS_ERROR)
    THEN
      // XTS state is transfered to higher up
      // --> check error and plausibility checks there
      _eState                             := E_PROGRESS.PROGRESS_ERROR;
    ELSIF (_XtsTransportState.State = E_XTS_TRANSPORT_STATE.TRANSPORT_INIT + E_PROGRESS.PROGRESS_DONE)
    THEN 
      _eState                             := E_PROGRESS.PROGRESS_PREPARE;
    END_IF
  //-----------------------------------------------------------------------------------------------------
  //-----------------------------------------------------------------------------------------------------
  E_PROGRESS.PROGRESS_PREPARE:
    _eResult                              := _ItfCollectors[_nInstance].Init(TRUE);
    IF (_eResult = E_PROGRESS.PROGRESS_ERROR)
    THEN
      memcpy(ADR(_nInstanceError), ADR(_nInstance), SIZEOF(_nInstance));

      _eState                             := E_PROGRESS.PROGRESS_ERROR;

      _stMsg.eType                        := E_MessageType.eMessageerror;
      _stMsg.eSubdevice                   := e_Subdevice.Application_Init;
      _stMsg.iErrorNumber                 := _nInstanceError;
      _stMsg.sText                        := concat(TO_STRING(_eState), ': ');
      _stMsg.sText                        := concat(_stMsg.sText, TO_STRING(_nInstanceError));
      f_MessageSet(_stMsg);

    ELSIF (_eResult = E_PROGRESS.PROGRESS_DONE)
    THEN
      _eState                             := E_PROGRESS.PROGRESS_STARTUP;
    END_IF
  //-----------------------------------------------------------------------------------------------------
  //-----------------------------------------------------------------------------------------------------
  E_PROGRESS.PROGRESS_STARTUP:
    IF (_nInstance < E_INSTANCE.INSTANCE_MAX-1)
    THEN
      _nInstance                          := _nInstance + 1;
      _eState                             := E_PROGRESS.PROGRESS_PREPARE;
    ELSE
      _eState                             := E_PROGRESS.PROGRESS_CHECK;
    END_IF
  //-----------------------------------------------------------------------------------------------------
  //-----------------------------------------------------------------------------------------------------
  E_PROGRESS.PROGRESS_CHECK:
    IF (_XtsTransportState.GroupInfo.GroupError)
    THEN
      _eState                             := E_PROGRESS.PROGRESS_ERROR;

      _stMsg.eType                        := E_MessageType.eMessageerror;
      _stMsg.eSubdevice                   := e_Subdevice.Application_Init;
      _stMsg.iErrorNumber                 := 0;
      _stMsg.sText                        := concat(TO_STRING(_eState), ': GroupInfo.GroupError');
      f_MessageSet(_stMsg);
    ELSE
      IF NOT (_XtsTransportState.XpuInfo.AllPositionsValid)
      THEN
        _eState                           := E_PROGRESS.PROGRESS_ERROR;
  
        _stMsg.eType                      := E_MessageType.eMessageerror;
        _stMsg.eSubdevice                 := e_Subdevice.Application_Init;
        _stMsg.iErrorNumber               := 0;
        _stMsg.sText                      := concat(TO_STRING(_eState), ': XpuInfo.AllPositionsValid');
        f_MessageSet(_stMsg);

      ELSE
        IF (_XtsTransportState.XpuInfo.IdDetectionValid) OR
           (_XtsTransportState.XpuInfo.IdDetectionMode = 0)
        THEN
          _eState                         := E_PROGRESS.PROGRESS_WORKING;
        END_IF
      END_IF
    END_IF
  //-----------------------------------------------------------------------------------------------------
  //-----------------------------------------------------------------------------------------------------
  E_PROGRESS.PROGRESS_WORKING:
    _eState                               := E_PROGRESS.PROGRESS_DONE;

    IF (_MessageLevel > E_MessageType.eMessageError)
    THEN
      _stMsg.eType                        := E_MessageType.eMessageInfo;
      _stMsg.eSubdevice                   := e_Subdevice.Application_Init;
      _stMsg.iErrorNumber                 := 0;
      _stMsg.sText                        := concat(TO_STRING(_eState), ': ');
      f_MessageSet(_stMsg);
    END_IF
END_CASE
//-------------------------------------------------------------------------------------------------------
//-------------------------------------------------------------------------------------------------------
Init                                      := _eState;
END_METHOD

PROPERTY MessageLevel : e_MessageType
GET
MessageLevel := _MessageLevel;
END_GET
SET
_MessageLevel := MessageLevel;
END_SET
END_PROPERTY

PROPERTY State : REFERENCE TO ST_YARD_STATE
SET
_State ref= State;
END_SET
END_PROPERTY

PROPERTY TicketList : I_Process_LinkedList
SET
_ItfTicketList := TicketList;
END_SET
END_PROPERTY

